FUNCTION_BLOCK FB_ProductionTank EXTENDS FB_SFC_Cycle IMPLEMENTS ITF_FB_SFC_Cycle
VAR_INPUT
	eElementID		: E_Element_List;
	
	stTankValves				:	st_TankValves		;
	stLineSourceValves			:	st_LineSourceValves	;
	stTriBlenderSourceValves	:	st_LineSourceValves	;
	stLineTargetValves			:	st_LineTargetValves	;
	stfbTriBlenderTargetValves	:	st_LineTargetValves	;

	
	
	//valOutlet		: E_Pis_Name;//Comment?
	//valLine			: E_Pis_Name;//Comment?
	//valTriBlender	: E_Pis_Name;//Comment?
	//valDrain		: E_Pis_Name;//Comment?
	//valCIP			: E_Pis_Name;//Comment?
	
	valFilling				: E_Pis_Name;
	valFillWater			: E_Pis_Name;
	valFillWaterDrain		: E_Pis_Name;
	valDrainTapWater		: E_Pis_Name;
	
	eTank_Name				: E_Tank_Name;

	
	sens_TankTemp			: E_ASense_Name	;//Tenk temperature sensor ID
	
	valCW_In				:	E_Pis_Name	;//Valve to control tank temperature In
	valCW_Out				:	E_Pis_Name	;//Valve to control tank temperature Out (always at 100 open)
	
	//pumpEnum			:	E_Pump_List	;
	
END_VAR
VAR_OUTPUT
END_VAR
VAR
	sTank_Name			: STRING;
	refElement			: REFERENCE TO FB_Element;
	refState_Long		: REFERENCE TO E_Element_State_Long;
	eReq				: E_Request_List;		
	eProcess			: E_Element_Process;
	eStatus				: E_Element_State_Long; // for HMI only as status
	
	fbPis				: FB_Piston;	
	
	//stPis_FillWater			: REFERENCE TO ST_Piston;
	//stPis_FillWaterDrain		: REFERENCE TO ST_Piston;
	//stPis_DrainTapWater		: REFERENCE TO ST_Piston;
	
	stPis_CWIn				: REFERENCE TO ST_Piston;
	stPis_CWOut				: REFERENCE TO ST_Piston;
	
	bTestingMode	:	BOOL	;//For testing purposes, to be deleted 
	bMoveStep		:	BOOL	;//For testing purposes, to be deleted 
	
	Call_TON	:	TON	;//Call ton for double request same object
	bTON_Active	:	BOOL	;
	
	// Temperature process control
	pc_TempCntrl	: REFERENCE TO FB_ProcessControl	;
	st_TempCntrl	: REFERENCE TO ST_ProcessControl	;
	bCntrlTemp		: BOOL	;
	bRunCIP			: BOOL	;
	
	ref_fbTankSensors			: REFERENCE TO FB_TankSensors;
	stTank_Level				: ST_Tank_Level;

	//888888888888888888888888888888888888888888
	stProdParam		: ST_Production_Parameter;
	//888888888888888888888888888888888888888888
	tonStirrer_time: TON;
	rTest: REAL := 16;
	bStirrerDirectionPositive: BOOL;
	
	delta_Tank_Volume		: REAL;
	memo_Tank_Level_start	: REAL;
	bRunOffline: BOOL;
	
	event_state_Update: INT;
	event_state_Update_sum: INT;
	event_state_Update_sum_last: INT;
	fbEvent_echo: FB_Event_echo;
	memo_Production_Storage_Mode: BOOL;
	memo_CIP_Pump_linked: BOOL;
	
	bStateUpdate_Available_HMI	: BOOL;

	
	
	fbFilling				: FB_Filling;		
	eFilling_State			: E_Filling_State;

END_VAR
VAR_IN_OUT

	fbTarget				: FB_Tank_Target;
	fbLineSource			: FB_Line_Source;
	fbLineTarget			: FB_Line_Target;
	fbTriBlenderSource		: FB_Line_Source;
	fbTriBlenderTarget		: FB_Line_Target;
	
	fbInterConnection_TriB	: FB_InterConnection;
	fbInterConnection_ProL	: FB_InterConnection;
	

	fb_PumpLine				: FB_Pump;
	fb_PumpTriBlender		: FB_Pump;
	fb_Stirrer				: FB_Pump;
END_VAR

act_GetReference();
act_Oper();
act_Call_Interface(); //There is no need to Call block if it comes from the outside
act_TempCntrl();
act_ExpirationTime();
act_Filling();

CASE eTank_Name OF
	E_Tank_Name.T1: sTank_Name:='Production Tank-T1';
	E_Tank_Name.T2: sTank_Name:='Production Tank-T2';
	E_Tank_Name.T3: sTank_Name:='Production Tank-T3';
	E_Tank_Name.T4: sTank_Name:='Production Tank-T4';
END_CASE

IF bTestingMode THEN;
	IF bMoveStep THEN;
		bMoveStep:=FALSE; 
	END_IF	
ELSE;
	bMoveStep:=TRUE; 
END_IF


IF stProdParam.bGetRecipe THEN;
	stProdParam.bGetRecipe:=FALSE;
	mGet_Recipe(indexRecipe:=stProdParam.hmiRecipeIndex+1);
END_IF
CASE eElementID	OF 
	E_Element_List.eTank_1,E_Element_List.eTank_2:;
		stProdParam.listRecipe:=g_Prod.listRecipe_Marinade;
	E_Element_List.eTank_3,E_Element_List.eTank_4:;
  		stProdParam.listRecipe:=g_Prod.listRecipe_Color;
END_CASE

stProdParam.timeRemainToStart:=mTimeRemainToStart();
stProdParam.timeProductionDuration:=mTimeProductionDuration();
refElement.ProdStatus:=stProdParam.eStatus;


IF refElement.m_Get_InterConnection()=E_InterConnection.NotConnected 
AND bReady
THEN;
	IF NOT bStateUpdate_Available_HMI THEN;
		refElement.fbEvent_echo.event();
		bStateUpdate_Available_HMI:=TRUE;
	END_IF	
ELSE; 
	IF bStateUpdate_Available_HMI THEN;
		refElement.fbEvent_echo.event();
		bStateUpdate_Available_HMI:=FALSE;
	END_IF
END_IF

m_Stirrer();
m_HMI();

ACTION _aCheck_Condition_Prod_End_active:
bStepDone:=FALSE;
IF fbInterConnection_ProL.bAvalableToDisconnect 
AND stProdParam.eStatus=E_Prod_Status.Active
THEN;
	bStepDone:=TRUE;
END_IF
END_ACTION

ACTION _aCheck_Condition_Product_active:
bStepDone:=FALSE;
IF fbInterConnection_ProL.bAvalableToConnect 
AND stProdParam.eStatus=E_Prod_Status.Active
THEN;
	bStepDone:=TRUE;
END_IF
END_ACTION

ACTION _aCheck_Condition_TriB_1_active_1:
bStepDone:=FALSE;
IF fbInterConnection_TriB.bAvalableToConnect
AND stProdParam.eStatus=E_Prod_Status.Active
AND m_Get_TriBlender_Clean()
THEN;
	bStepDone:=TRUE;
END_IF
END_ACTION

ACTION _aCheck_Condition_TriB_2_active:
bStepDone:=FALSE;
IF fbInterConnection_TriB.bAvalableToConnect 
AND stProdParam.eStatus=E_Prod_Status.Active
AND m_Get_TriBlender_Clean()
THEN;
	bStepDone:=TRUE;
END_IF
END_ACTION

ACTION _aClose_01_active:
bStepDone:=FALSE;
IF fbTarget.m_CheckStatus(eReqStatus:=E_Tank_Target.eClose) THEN;
	bStepDone:=TRUE;
END_IF
END_ACTION

ACTION _aClose_01_entry:
fbTarget.m_Run(eReqProc:=E_Tank_Target.eClose);
END_ACTION

ACTION _aClose_2_active:
bStepDone:=FALSE;
IF fbTarget.m_CheckStatus(eReqStatus:=E_Tank_Target.eClose) THEN;
	bStepDone:=TRUE;
END_IF
END_ACTION

ACTION _aClose_2_entry:
fbTarget.m_Run(eReqProc:=E_Tank_Target.eClose);
END_ACTION

ACTION _aClose_4_active:
bStepDone:=FALSE;
IF fbTarget.m_CheckStatus(eReqStatus:=E_Tank_Target.eClose) THEN;
	bStepDone:=TRUE;
END_IF
END_ACTION

ACTION _aClose_4_entry:
fbTarget.m_Run(eReqProc:=E_Tank_Target.eClose);
END_ACTION

ACTION _aClose_Drain_val_active:
//bStepDone:=FALSE;
IF fbTarget.m_CheckStatus(eReqStatus:=E_Tank_Target.eOpen) THEN;
(*ELSE
	fbTarget.m_Run(eReqProc:=E_Tank_Target.eOpen);*)
	bTON_Active:=TRUE;
END_IF
IF Call_TON.Q THEN
	bStepDone:=TRUE;
END_IF
END_ACTION

ACTION _aClose_Drain_val_entry:
bStepDone:=FALSE;
fbTarget.m_Run(eReqProc:=E_Tank_Target.eOpen);
bTON_Active:=FALSE;
END_ACTION

ACTION _aClose_Tank_active:
bStepDone:=FALSE;
IF fbTarget.m_CheckStatus(eReqStatus:=E_Tank_Target.eClose_DrainPipe) THEN;
	bStepDone:=TRUE;
END_IF
END_ACTION

ACTION _aClose_Tank_entry:
fbTarget.m_Run(eReqProc:=E_Tank_Target.eClose_DrainPipe);
END_ACTION

ACTION _aCollect_From_Prod_Line_active:
bStepDone:=FALSE;
delta_Tank_Volume:=ref_fbTankSensors.act_Volume-memo_Tank_Level_start;
IF FALSE 
OR delta_Tank_Volume>=stProdParam.stRecipe.Weight_to_Collect
OR Collect_From_Prod_Line.t>=T#40S
THEN;
	bStepDone:=TRUE;
END_IF
END_ACTION

ACTION _aCollect_From_TriB_Line_active:
bStepDone:=FALSE;
delta_Tank_Volume:=ref_fbTankSensors.act_Volume-memo_Tank_Level_start;
IF FALSE 
OR delta_Tank_Volume>=stProdParam.stRecipe.Weight_to_Collect
OR Collect_From_TriB_Line.t>=T#40S
THEN;
	bStepDone:=TRUE;
END_IF
END_ACTION

ACTION _aConn_Line_Source_TankA_active:
bStepDone:=FALSE;
IF fbLineSource.m_CheckStatus(eReqStatus:=E_Line_Source.eTank_A) THEN;
	bStepDone:=TRUE;
END_IF
END_ACTION

ACTION _aConn_Line_Source_TankA_entry:
fbLineSource.m_Run(eReqProc:=E_Line_Source.eTank_A);
END_ACTION

ACTION _aConn_Line_Source_TankB_active:
bStepDone:=FALSE;
IF fbLineSource.m_CheckStatus(eReqStatus:=E_Line_Source.eTank_B) THEN;
	bStepDone:=TRUE;
END_IF
END_ACTION

ACTION _aConn_Line_Source_TankB_entry:
fbLineSource.m_Run(eReqProc:=E_Line_Source.eTank_B);
END_ACTION

ACTION _aConn_Line_Target_TankA_active:
bStepDone:=FALSE;
IF fbLineTarget.m_CheckStatus(eReqStatus:=E_Line_Target.eTank_A) THEN;
	bTON_Active:=TRUE;
END_IF
IF Call_TON.Q THEN
	bStepDone:=TRUE;
END_IF
END_ACTION

ACTION _aConn_Line_Target_TankA_entry:
fbLineTarget.m_Run(eReqProc:=E_Line_Target.eTank_A);
bTON_Active:=FALSE;
END_ACTION

ACTION _aConn_Line_Target_TankB_active:
bStepDone:=FALSE;
IF fbLineTarget.m_CheckStatus(eReqStatus:=E_Line_Target.eTank_B) THEN;
	bTON_Active:=TRUE;
END_IF
IF Call_TON.Q THEN
	bStepDone:=TRUE;
END_IF
END_ACTION

ACTION _aConn_Line_Target_TankB_entry:
fbLineTarget.m_Run(eReqProc:=E_Line_Target.eTank_B);
bTON_Active:=FALSE;
END_ACTION

ACTION _aConn_Tank_active:
bStepDone:=FALSE;
IF fbTriBlenderSource.m_CheckStatus(eReqStatus:=E_Line_Source.eFillWater) 
//AND fbPis.m_CheckByRecipe(stPis:=stPis_FillWaterDrain, req:=E_Piston_Recipe_State.Release) 
THEN;
	bStepDone:=TRUE;
END_IF
END_ACTION

ACTION _aConn_Tank_entry:
fbTriBlenderSource.m_Run(eReqProc:=E_Line_Source.eFillWater);
//fbPis.m_SetByRecipe(stPis:=stPis_FillWaterDrain, req:=E_Piston_Recipe_State.Release);
END_ACTION

ACTION _aConn_Tri_Drain_active:
bStepDone:=FALSE;
IF fbTriBlenderTarget.m_CheckStatus(eReqStatus:=E_Line_Target.eDrain) THEN;
	bStepDone:=TRUE;
END_IF
END_ACTION

ACTION _aConn_Tri_Drain_entry:
fbTriBlenderTarget.m_Run(eReqProc:=E_Line_Target.eDrain);
END_ACTION

ACTION _aConn_Tri_TankA_2_active:
bStepDone:=FALSE;
IF fbTriBlenderSource.m_CheckStatus(eReqStatus:=E_Line_Source.eTank_A) THEN;
	bStepDone:=TRUE;
END_IF
END_ACTION

ACTION _aConn_Tri_TankA_2_entry:
fbTriBlenderSource.m_Run(eReqProc:=E_Line_Source.eTank_A);
END_ACTION

ACTION _aConn_Tri_TankB_2_active:
bStepDone:=FALSE;
IF fbTriBlenderSource.m_CheckStatus(eReqStatus:=E_Line_Source.eTank_B) THEN;
	bStepDone:=TRUE;
END_IF
END_ACTION

ACTION _aConn_Tri_TankB_2_entry:
fbTriBlenderSource.m_Run(eReqProc:=E_Line_Source.eTank_B);
END_ACTION

ACTION _aConn_Tri_TapWater_active:
bStepDone:=FALSE;
IF fbTriBlenderSource.m_CheckStatus(eReqStatus:=E_Line_Source.eTapWater) 
//AND fbPis.m_CheckByRecipe(stPis:=stPis_DrainTapWater, req:=E_Piston_Recipe_State.Release) 
THEN;
	bTON_Active:=TRUE;
END_IF
IF Call_TON.Q THEN
	bStepDone:=TRUE;
END_IF
END_ACTION

ACTION _aConn_Tri_TapWater_entry:
fbTriBlenderSource.m_Run(eReqProc:=E_Line_Source.eTapWater);
//fbPis.m_SetByRecipe(stPis:=stPis_DrainTapWater, req:=E_Piston_Recipe_State.Release);
bTON_Active:=FALSE;
END_ACTION

ACTION _aConn_Tri_ToTankA_1_active:
bStepDone:=FALSE;
IF fbTriBlenderTarget.m_CheckStatus(eReqStatus:=E_Line_Target.eTank_A) THEN;
	bStepDone:=TRUE;
END_IF
END_ACTION

ACTION _aConn_Tri_ToTankA_1_entry:
fbTriBlenderTarget.m_Run(eReqProc:=E_Line_Target.eTank_A);
END_ACTION

ACTION _aConn_Tri_ToTankA_2_active:
bStepDone:=FALSE;
IF fbTriBlenderTarget.m_CheckStatus(eReqStatus:=E_Line_Target.eTank_A) THEN;
	bStepDone:=TRUE;
END_IF
END_ACTION

ACTION _aConn_Tri_ToTankA_2_entry:
fbTriBlenderTarget.m_Run(eReqProc:=E_Line_Target.eTank_A);
END_ACTION

ACTION _aConn_Tri_ToTankB_1_active:
bStepDone:=FALSE;
IF fbTriBlenderTarget.m_CheckStatus(eReqStatus:=E_Line_Target.eTank_B) THEN;
	bStepDone:=TRUE;
END_IF
END_ACTION

ACTION _aConn_Tri_ToTankB_1_entry:
fbTriBlenderTarget.m_Run(eReqProc:=E_Line_Target.eTank_B);
END_ACTION

ACTION _aConn_Tri_ToTankB_2_active:
bStepDone:=FALSE;
IF fbTriBlenderTarget.m_CheckStatus(eReqStatus:=E_Line_Target.eTank_B) THEN;
	bStepDone:=TRUE;
END_IF
END_ACTION

ACTION _aConn_Tri_ToTankB_2_entry:
fbTriBlenderTarget.m_Run(eReqProc:=E_Line_Target.eTank_B);
END_ACTION

ACTION _aConn_TriB_Color_active_1:
bStepDone:=FALSE;
IF fbTriBlender_Select.m_CheckStatus(eReqStatus:=E_TriBlenderSelect.eColor) THEN;
	bStepDone:=TRUE;
END_IF
END_ACTION

ACTION _aConn_TriB_Color_entry_1:
fbTriBlender_Select.m_Set_Request(eSetReg:=E_TriBlenderSelect.eColor);
END_ACTION

ACTION _aConn_TriB_Marinade_active_1:
bStepDone:=FALSE;
IF fbTriBlender_Select.m_CheckStatus(eReqStatus:=E_TriBlenderSelect.eMarinade) THEN;
	bStepDone:=TRUE;
END_IF
END_ACTION

ACTION _aConn_TriB_Marinade_entry_1:
fbTriBlender_Select.m_Set_Request(eSetReg:=E_TriBlenderSelect.eMarinade);
END_ACTION

ACTION _aDis_Conn_Tank_active:
bStepDone:=FALSE;
IF fbTriBlenderSource.m_CheckStatus(eReqStatus:=E_Line_Source.eClose) 
AND fbTriBlenderTarget.m_CheckStatus(eReqStatus:=E_Line_Target.eDrain) 
THEN;
	bStepDone:=TRUE;
END_IF
END_ACTION

ACTION _aDis_Conn_Tank_entry:
fbTriBlenderSource.m_Run(eReqProc:=E_Line_Source.eClose);
fbTriBlenderTarget.m_Run(eReqProc:=E_Line_Target.eDrain);
END_ACTION

ACTION _aDisconn_Tri_Tank_active:
bStepDone:=FALSE;
IF fbTriBlenderSource.m_CheckStatus(eReqStatus:=E_Line_Source.eClose) THEN;
	bTON_Active:=TRUE;
END_IF
IF Call_TON.Q THEN
	bStepDone:=TRUE;
END_IF
END_ACTION

ACTION _aDisconn_Tri_Tank_entry:
fbTriBlenderSource.m_Run(eReqProc:=E_Line_Source.eClose);
bTON_Active:=FALSE;
END_ACTION

ACTION _aDisconnect_TapWater_02_active:
bStepDone:=FALSE;
IF fbTriBlenderSource.m_CheckStatus(eReqStatus:=E_Line_Source.eDrain) THEN;
	bStepDone:=TRUE;
END_IF
END_ACTION

ACTION _aDisconnect_TapWater_02_entry:
fbTriBlenderSource.m_Run(eReqProc:=E_Line_Source.eDrain);
END_ACTION

ACTION _aDissolving_entry:
bDisolvingProcess_Done:=FALSE;
bDisolvingProcess_Active:=FALSE;
END_ACTION

ACTION _aDissolving_Proc_active:
bStepDone:=FALSE;

IF bDisolvingProcess_Done 
//AND fbDissolving.bD
THEN;
	
END_IF
END_ACTION

ACTION _aDissolving_Proc_entry:

bDisolvingProcess_Active:=TRUE;
fbDissolving.mRun();
END_ACTION

ACTION _aDissolving_Proc_exit:
bDisolvingProcess_Done:=FALSE;
bDisolvingProcess_Active:=FALSE;
END_ACTION

ACTION _aDone_entry:
eProcess:=E_Element_Process.eNone;
eReq:=E_Request_List.eNone;
bRun:=FALSE;
bDone:=TRUE;
END_ACTION

ACTION _aDrain_All_Marinade_Lines_active:
bStepDone:=FALSE;
IF TRUE
//AND fbTarget.m_CheckStatus(eReqStatus:=E_Tank_Target.eClose_DrainPipe) 
AND fbTriBlenderSource.m_CheckStatus(eReqStatus:=E_Line_Source.eDrain)
AND fbTriBlenderTarget.m_CheckStatus(eReqStatus:=E_Line_Target.eDrain)
AND fbTriBlender_Select.m_CheckStatus(eReqStatus:=E_TriBlenderSelect.eDrain)
AND TRUE
AND TRUE
THEN;
	bStepDone:=TRUE;
END_IF
END_ACTION

ACTION _aDrain_All_Marinade_Lines_entry:
//fbTarget.m_Run(eReqProc:=E_Tank_Target.eClose_DrainPipe);
fbTriBlenderSource.m_Run(eReqProc:=E_Line_Source.eDrain);
fbTriBlenderTarget.m_Run(eReqProc:=E_Line_Target.eDrain);
fbTriBlender_Select.m_Set_Request(eSetReg:=E_TriBlenderSelect.eDrain);
END_ACTION

ACTION _aDrain_Pipe_active:
bStepDone:=FALSE;
IF fbTarget.m_CheckStatus(eReqStatus:=E_Tank_Target.eClose_DrainPipe) THEN;
	bTON_Active:=TRUE;
END_IF
IF Call_TON.Q THEN
	bStepDone:=TRUE;
END_IF
END_ACTION

ACTION _aDrain_Pipe_Close_active:
bStepDone:=FALSE;
IF fbTarget.m_CheckStatus(eReqStatus:=E_Tank_Target.eClose) THEN;
	bStepDone:=TRUE;
END_IF
END_ACTION

ACTION _aDrain_Pipe_Close_entry:
fbTarget.m_Run(eReqProc:=E_Tank_Target.eClose);
END_ACTION

ACTION _aDrain_Pipe_entry:
fbTarget.m_Run(eReqProc:=E_Tank_Target.eClose_DrainPipe);
bTON_Active:=FALSE;
END_ACTION

ACTION _aDrain_Production_Line_active:
bStepDone:=FALSE;
IF TRUE
AND fbTarget.m_CheckStatus(eReqStatus:=E_Tank_Target.eClose_DrainPipe) 
AND fbLineSource.m_CheckStatus(eReqStatus:=E_Line_Source.eDrain)
AND fbLineTarget.m_CheckStatus(eReqStatus:=E_Line_Target.eDrain)
AND TRUE
THEN;
	bStepDone:=TRUE;
END_IF
END_ACTION

ACTION _aDrain_Production_Line_entry:
fbTarget.m_Run(eReqProc:=E_Tank_Target.eClose_DrainPipe);
fbLineSource.m_Run(eReqProc:=E_Line_Source.eDrain);
fbLineTarget.m_Run(eReqProc:=E_Line_Target.eDrain);
END_ACTION

ACTION _aDrain_Tri_Line_active:
bStepDone:=FALSE;
IF fbTriBlenderTarget.m_CheckStatus(eReqStatus:=E_Line_Target.eDrain) THEN;
	bStepDone:=TRUE;
END_IF
END_ACTION

ACTION _aDrain_Tri_Line_entry:
fbTriBlenderTarget.m_Run(eReqProc:=E_Line_Target.eDrain);
END_ACTION

ACTION _aDrain_Tri_ToDrain_active:
bStepDone:=FALSE;
IF fbTriBlenderTarget.m_CheckStatus(eReqStatus:=E_Line_Target.eDrain) THEN;
	bTON_Active:=TRUE;
END_IF
IF Call_TON.Q THEN
	bStepDone:=TRUE;
END_IF

(*
delta_Tank_Volume:=ref_fbTankSensors.act_Volume-memo_Tank_Level_start;
IF bStepDone
AND  
AND (delta_Tank_Volume>=stProdParam.stRecipe.Weight_to_Drain
	OR Drain_Tri_ToDrain.t>=T#30S)
THEN;
	//bStepDone:=TRUE;
ELSE;
	bStepDone:=FALSE;
END_IF
*)
END_ACTION

ACTION _aDrain_Tri_ToDrain_entry:
fbTriBlenderTarget.m_Run(eReqProc:=E_Line_Target.eDrain);
bTON_Active:=FALSE;
END_ACTION

ACTION _aDrain_Tri_ToTankA_active:
bStepDone:=FALSE;
IF fbTriBlenderTarget.m_CheckStatus(eReqStatus:=E_Line_Target.eTank_A) THEN;
	bTON_Active:=TRUE;
END_IF
IF Call_TON.Q THEN
	bStepDone:=TRUE;
END_IF
END_ACTION

ACTION _aDrain_Tri_ToTankA_entry:
fbTriBlenderTarget.m_Run(eReqProc:=E_Line_Target.eTank_A);
bTON_Active:=FALSE;
END_ACTION

ACTION _aDrain_Tri_ToTankB_active:
bStepDone:=FALSE;
IF fbTriBlenderTarget.m_CheckStatus(eReqStatus:=E_Line_Target.eTank_B) THEN;
	bTON_Active:=TRUE;
END_IF
IF Call_TON.Q THEN
	bStepDone:=TRUE;
END_IF
END_ACTION

ACTION _aDrain_Tri_ToTankB_entry:
fbTriBlenderTarget.m_Run(eReqProc:=E_Line_Target.eTank_B);
bTON_Active:=FALSE;
END_ACTION

ACTION _aDrain_Trib_Line_01_active:
bStepDone:=FALSE;
IF fbTriBlender_Select.m_CheckStatus(eReqStatus:=E_TriBlenderSelect.eDrain) THEN;
	bStepDone:=TRUE;
END_IF
END_ACTION

ACTION _aDrain_Trib_Line_01_entry:
fbTriBlender_Select.m_Set_Request(eSetReg:=E_TriBlenderSelect.eDrain);
END_ACTION

ACTION _aDrain_Trib_Line_02_active:
bStepDone:=FALSE;
IF fbTriBlender_Select.m_CheckStatus(eReqStatus:=E_TriBlenderSelect.eDrain)
OR fbTriBlender_Select.m_CheckStatus(eReqStatus:=E_TriBlenderSelect.eMarinade) THEN;//marinade =>> drain time finish
	bStepDone:=TRUE;
END_IF
END_ACTION

ACTION _aDrain_Trib_Line_02_entry:
fbTriBlender_Select.m_Set_Request(eSetReg:=E_TriBlenderSelect.eDrain);
END_ACTION

ACTION _aDraining_Time_active:
bStepDone:=FALSE;
IF stTank_Level.e_state=E_Tank_Level.eEmpty THEN;
	bStepDone:=TRUE;
END_IF
END_ACTION

ACTION _aDrainOpen_01_active:
bStepDone:=FALSE;
IF fbTarget.m_CheckStatus(eReqStatus:=E_Tank_Target.eDrain) THEN;
	bStepDone:=TRUE;
END_IF
END_ACTION

ACTION _aDrainOpen_01_entry:
fbTarget.m_Run(eReqProc:=E_Tank_Target.eDrain);
END_ACTION

ACTION _aDriin_Tank_active:
bStepDone:=FALSE;
IF stTank_Level.e_state=E_Tank_Level.eEmpty THEN;
	bStepDone:=TRUE;
END_IF
END_ACTION

ACTION _aDriin_Tank_entry:
fbTarget.m_Run(eReqProc:=E_Tank_Target.eDrain);
END_ACTION

ACTION _aInit_Base_active:
bStepDone:=FALSE;
IF TRUE
AND refState_Long<>E_Element_State_Long.eProduction
AND fbTarget.m_CheckStatus(eReqStatus:=E_Tank_Target.eClose_DrainPipe) 
AND TRUE
THEN;
	bStepDone:=TRUE;
ELSIF refState_Long=E_Element_State_Long.eProduction THEN;
	bStepDone:=TRUE;
END_IF
END_ACTION

ACTION _aInit_Base_entry:
IF refState_Long<>E_Element_State_Long.eProduction THEN;	
	fb_PumpLine.m_Stop();
	fbTarget.m_Run(eReqProc:=E_Tank_Target.eClose_DrainPipe);
END_IF
END_ACTION

ACTION _aInit_Production_Line_active:
bStepDone:=FALSE;
IF TRUE
AND refState_Long<>E_Element_State_Long.eProduction
AND fbTarget.m_CheckStatus(eReqStatus:=E_Tank_Target.eClose_DrainPipe) 
AND fbLineSource.m_CheckStatus(eReqStatus:=E_Line_Source.eDrain)
AND fbLineTarget.m_CheckStatus(eReqStatus:=E_Line_Target.eDrain)
AND (NOT fbInterConnection_ProL.bActive)
AND TRUE
THEN;
	bStepDone:=TRUE;
ELSIF refState_Long=E_Element_State_Long.eProduction THEN;
	bStepDone:=TRUE;
END_IF
END_ACTION

ACTION _aInit_Production_Line_entry:
IF refState_Long<>E_Element_State_Long.eProduction THEN;	
	fb_PumpLine.m_Stop();
	fbTarget.m_Run(eReqProc:=E_Tank_Target.eClose_DrainPipe);
	fbLineSource.m_Run(eReqProc:=E_Line_Source.eDrain);
	fbLineTarget.m_Run(eReqProc:=E_Line_Target.eDrain);
	fbInterConnection_ProL.reqDisconnect:=TRUE;
END_IF
END_ACTION

ACTION _aInit_Tank_active:
SFCReset:=FALSE;
END_ACTION

ACTION _aInit_Tank_exit:
IF eProcess=E_Element_Process.eFill_Water THEN;
	mClearProduction(state:=E_Element_State_Long.eOff);
END_IF

eProcess:=E_Element_Process.eNone;
eReq:=E_Request_List.eNone;
memo_Production_Storage_Mode:=FALSE;
END_ACTION

ACTION _aInit_TriBlender_Line_active:
bStepDone:=FALSE;
IF TRUE
AND fbTarget.m_CheckStatus(eReqStatus:=E_Tank_Target.eClose_DrainPipe) 
AND fbTriBlenderSource.m_CheckStatus(eReqStatus:=E_Line_Source.eDrain)
AND fbTriBlenderTarget.m_CheckStatus(eReqStatus:=E_Line_Target.eDrain)
AND fbTriBlender_Select.m_CheckStatus(eReqStatus:=E_TriBlenderSelect.eDrain)
AND (NOT fbInterConnection_TriB.bActive)
AND TRUE
THEN;
	bStepDone:=TRUE;
END_IF
END_ACTION

ACTION _aInit_TriBlender_Line_entry:
fb_PumpTriBlender.m_Stop();
fbTarget.m_Run(eReqProc:=E_Tank_Target.eClose_DrainPipe);
fbTriBlenderSource.m_Run(eReqProc:=E_Line_Source.eDrain);
fbTriBlenderTarget.m_Run(eReqProc:=E_Line_Target.eDrain);
fbTriBlender_Select.m_Set_Request(eSetReg:=E_TriBlenderSelect.eDrain);
fbInterConnection_TriB.reqDisconnect:=TRUE;
fbDissolving.mResetCycle();
END_ACTION

ACTION _aInterConnect_Prod_active:
bStepDone:=FALSE;
IF fbInterConnection_ProL.bActive THEN;
	bStepDone:=TRUE;
END_IF
END_ACTION

ACTION _aInterConnect_Prod_Dis_active:
bStepDone:=FALSE;
IF NOT fbInterConnection_ProL.bActive THEN;
	bStepDone:=TRUE;
END_IF
END_ACTION

ACTION _aInterConnect_Prod_Dis_entry:
fbInterConnection_ProL.reqDisconnect:=TRUE;
END_ACTION

ACTION _aInterConnect_Prod_entry:
fbInterConnection_ProL.reqConnect:=TRUE;

IF trn_Tank_Marinade THEN;
	//fbElement[E_Element_List.eTriBlender_Marinada].m_Set_Dissolveng_active_memo();
ELSIF trn_Tank_Color THEN;
	//fbElement[E_Element_List.eTriBlender_Color].m_Set_Dissolveng_active_memo();
END_IF
END_ACTION

ACTION _aInterConnect_TriB_1_active:
bStepDone:=FALSE;
IF fbInterConnection_TriB.bActive THEN;
	bStepDone:=TRUE;
END_IF
END_ACTION

ACTION _aInterConnect_TriB_1_entry:
fbInterConnection_TriB.reqConnect:=TRUE;
END_ACTION

ACTION _aInterConnect_TriB_2_active:
bStepDone:=FALSE;
IF fbInterConnection_TriB.bActive THEN;
	bStepDone:=TRUE;
	
	refElement.m_Set_Dissolveng_active_memo();
	IF trn_Tank_Marinade THEN;
		fbElement[E_Element_List.eTriBlender_Marinada].m_Set_Dissolveng_active_memo();
	ELSIF trn_Tank_Color THEN;
		fbElement[E_Element_List.eTriBlender_Color].m_Set_Dissolveng_active_memo();
	ELSE;
		bStepDone:=FALSE;
	END_IF	
	
END_IF
END_ACTION

ACTION _aInterConnect_TriB_2_entry:
fbInterConnection_TriB.reqConnect:=TRUE;
END_ACTION

ACTION _aInterConnect_TriB_Dis_1_active:
bStepDone:=FALSE;
IF NOT fbInterConnection_TriB.bActive THEN;
	bStepDone:=TRUE;
END_IF
END_ACTION

ACTION _aInterConnect_TriB_Dis_1_entry:
fbInterConnection_TriB.reqDisconnect:=TRUE;
END_ACTION

ACTION _aInterConnect_TriB_Dis_2_active:
bStepDone:=FALSE;
IF NOT fbInterConnection_TriB.bActive THEN;
	bStepDone:=TRUE;
END_IF
END_ACTION

ACTION _aInterConnect_TriB_Dis_2_entry:
fbInterConnection_TriB.reqDisconnect:=TRUE;
END_ACTION

ACTION _aLineSource_Close_active:
bStepDone:=FALSE;
IF fbLineSource.m_CheckStatus(eReqStatus:=E_Line_Source.eClose) 
THEN;
	bStepDone:=TRUE;
END_IF
END_ACTION

ACTION _aLineSource_Close_entry:
fbLineSource.m_Run(eReqProc:=E_Line_Source.eClose);
END_ACTION

ACTION _aLineSource_TapWater_active:
bStepDone:=FALSE;
IF fbLineSource.m_CheckStatus(eReqStatus:=E_Line_Source.eTapWater) 
THEN;
	bStepDone:=TRUE;
END_IF
END_ACTION

ACTION _aLineSource_TapWater_entry:
fbLineSource.m_Run(eReqProc:=E_Line_Source.eTapWater);
bTON_Active:=FALSE;
END_ACTION

ACTION _aLineTarget_Drain_1_active:
bStepDone:=FALSE;
IF fbLineTarget.m_CheckStatus(eReqStatus:=E_Line_Target.eDrain) THEN;
	bStepDone:=TRUE;
END_IF
END_ACTION

ACTION _aLineTarget_Drain_1_entry:
fbLineTarget.m_Run(eReqProc:=E_Line_Target.eDrain);
END_ACTION

ACTION _aLineTarget_Drain_2_active:
bStepDone:=FALSE;
IF fbLineTarget.m_CheckStatus(eReqStatus:=E_Line_Target.eDrain) THEN;
	bTON_Active:=TRUE;
END_IF
IF Call_TON.Q THEN
	bStepDone:=TRUE;
END_IF
END_ACTION

ACTION _aLineTarget_Drain_2_entry:
fbLineTarget.m_Run(eReqProc:=E_Line_Target.eDrain);
bTON_Active:=FALSE;
END_ACTION

ACTION _aLineTarget_TankA_active:
bStepDone:=FALSE;
IF fbLineTarget.m_CheckStatus(eReqStatus:=E_Line_Target.eTank_A) THEN;
	bTON_Active:=TRUE;
END_IF
IF Call_TON.Q THEN
	bStepDone:=TRUE;
END_IF
END_ACTION

ACTION _aLineTarget_TankA_entry:
fbLineTarget.m_Run(eReqProc:=E_Line_Target.eTank_A);
bTON_Active:=FALSE;
END_ACTION

ACTION _aLineTarget_TankB_active:
bStepDone:=FALSE;
IF fbLineTarget.m_CheckStatus(eReqStatus:=E_Line_Target.eTank_B) THEN;
	bTON_Active:=TRUE;
END_IF
IF Call_TON.Q THEN
	bStepDone:=TRUE;
END_IF
END_ACTION

ACTION _aLineTarget_TankB_entry:
fbLineTarget.m_Run(eReqProc:=E_Line_Target.eTank_B);
bTON_Active:=FALSE;
END_ACTION

ACTION _aOpen_Drain_Pipe_active:
bStepDone:=FALSE;
IF fbTarget.m_CheckStatus(eReqStatus:=E_Tank_Target.eClose_DrainPipe) THEN;
	bStepDone:=TRUE;
END_IF
END_ACTION

ACTION _aOpen_Drain_Pipe_entry:
fbTarget.m_Run(eReqProc:=E_Tank_Target.eClose_DrainPipe);
END_ACTION

ACTION _aPumpLine_Auto_1_entry:
//fb_PumpLine.m_Auto();
END_ACTION

ACTION _aPumpLine_Start_1_active:

END_ACTION

ACTION _aPumpLine_Start_1_entry:
fb_PumpLine.m_Run(RPM:=stProdParam.stRecipe.FlowRate_Production);
END_ACTION

ACTION _aPumpLine_Start_2_entry:
fb_PumpLine.m_Run(RPM:=stProdParam.stRecipe.FlowRate_Production);
memo_Tank_Level_start:=ref_fbTankSensors.act_Volume;
END_ACTION

ACTION _aPumpLine_Stop_1_entry:
fb_PumpLine.m_Stop();
END_ACTION

ACTION _aPumpLine_Stop_2_entry:

IF trn_Tank_Marinade THEN;
	fb_PumpLine.m_Stop();
END_IF
END_ACTION

ACTION _aPumpLine_Stop_3_entry:
fb_PumpLine.m_Stop();
END_ACTION

ACTION _aPumpLine_Stop_4_entry:
fb_PumpLine.m_Stop();
END_ACTION

ACTION _aReady_active:


CASE refElement.eState_Long OF
	E_Element_State_Long.eOff,E_Element_State_Long.eStandby:;
			IF eReq=E_Request_List.eDrain THEN;
				eProcess:=E_Element_Process.eDrain;
			END_IF

	E_Element_State_Long.eCIP_5_Done:;
			IF eReq=E_Request_List.eWaterPrepare THEN;
				eProcess:=E_Element_Process.eFill_Water;
			END_IF	
			
	E_Element_State_Long.eWaterReady:;
			IF eReq=E_Request_List.eDissolve THEN;
				eProcess:=E_Element_Process.eDissolving;
			END_IF	
			IF eReq=E_Request_List.eFinish THEN;
				mClearProduction(state:=E_Element_State_Long.eStandby);
			END_IF
	E_Element_State_Long.eReady:;
			IF eReq=E_Request_List.eProduction THEN;
				eProcess:=E_Element_Process.eConnectionToLine;
			END_IF	
			IF eReq=E_Request_List.eFinish THEN;
				mClearProduction(state:=E_Element_State_Long.eStandby);
			END_IF			

	E_Element_State_Long.eProduction:;
			IF eReq=E_Request_List.eDisconnectTank THEN;
				eProcess:=E_Element_Process.eDisconnection;
			END_IF	
			
			IF fbInterConnection_ProL.bAvalableToDisconnect 
			AND m_Production_Run_Pump()
			THEN;
				IF memo_Production_Storage_Mode THEN;
					fb_PumpLine.m_Run(RPM:=stProdParam.stRecipe.FlowRate_Storage);
				ELSE;
					fb_PumpLine.m_Run(RPM:=stProdParam.stRecipe.FlowRate_Production);
				END_IF
				
			ELSE;
				fb_PumpLine.m_Stop();
			END_IF		

	E_Element_State_Long.eEmpty:;
			IF eReq=E_Request_List.eFinish THEN;
				mClearProduction(state:=E_Element_State_Long.eStandby);
			END_IF	

	E_Element_State_Long.eExpired:;
		CASE refElement.eState_Long_Expiered OF
			
			E_Element_State_Long.eProduction:;	
				IF eReq=E_Request_List.eDisconnectTank THEN;
					eProcess:=E_Element_Process.eDisconnection;
				END_IF
				
				IF fbInterConnection_ProL.bAvalableToDisconnect 
				AND m_Production_Run_Pump()
				THEN;
					IF memo_Production_Storage_Mode THEN;
						fb_PumpLine.m_Run(RPM:=stProdParam.stRecipe.FlowRate_Storage);
					ELSE;
						fb_PumpLine.m_Run(RPM:=stProdParam.stRecipe.FlowRate_Production);
					END_IF
					
				ELSE;
					fb_PumpLine.m_Stop();
				END_IF	
		ELSE
			IF eReq=E_Request_List.eFinish THEN;
				mClearProduction(state:=E_Element_State_Long.eStandby);
			END_IF			
		END_CASE
		
END_CASE
END_ACTION

ACTION _aReady_entry:

END_ACTION

ACTION _aReady_exit:
bRun:=TRUE;
bDone:=FALSE;
//bCntrlTemp:=TRUE;
END_ACTION

ACTION _aStart_TriPump_1_active:
bStepDone:=TRUE;
END_ACTION

ACTION _aStart_TriPump_1_entry:
fb_PumpTriBlender.m_Run(RPM:=stProdParam.stRecipe.FlowRate_WaterPushing);
END_ACTION

ACTION _aStart_TriPump_2_active:
bStepDone:=TRUE;
END_ACTION

ACTION _aStart_TriPump_2_entry:
fb_PumpTriBlender.m_Run(RPM:=stProdParam.stRecipe.FlowRate_WaterPushing);
END_ACTION

ACTION _aStart_TriPump_3_active:
bStepDone:=TRUE;
END_ACTION

ACTION _aStart_TriPump_3_entry:
fb_PumpTriBlender.m_Run(RPM:=stProdParam.stRecipe.FlowRate_WaterPushing);
memo_Tank_Level_start:=ref_fbTankSensors.act_Volume;
END_ACTION

ACTION _aState_Update_01_entry:
refState_Long:=E_Element_State_Long.eNotClean;
END_ACTION

ACTION _aState_Update_02_entry:
refState_Long:=E_Element_State_Long.eWaterReady;
END_ACTION

ACTION _aState_Update_03_entry:
refState_Long:=E_Element_State_Long.eReady;
END_ACTION

ACTION _aState_Update_04_entry:
refState_Long:=E_Element_State_Long.eProduction;
END_ACTION

ACTION _aState_Update_05_entry:
refState_Long:=E_Element_State_Long.eReady;
END_ACTION

ACTION _aStop_TriPump_1_active:
bStepDone:=TRUE;
END_ACTION

ACTION _aStop_TriPump_1_entry:
fb_PumpTriBlender.m_Stop();
END_ACTION

ACTION _aStop_TriPump_2_active:
bStepDone:=TRUE;
END_ACTION

ACTION _aStop_TriPump_2_entry:
fb_PumpTriBlender.m_Stop();
END_ACTION

ACTION _aStop_TriPump_3_active:
bStepDone:=TRUE;
END_ACTION

ACTION _aStop_TriPump_3_entry:
fb_PumpTriBlender.m_Stop();
END_ACTION

ACTION _aTank_Drain_active:
bStepDone:=FALSE;
IF fbTarget.m_CheckStatus(eReqStatus:=E_Tank_Target.eDrain) THEN;
	bTON_Active:=TRUE;
	
ELSIF Tank_Drain.t>=T#3S THEN; // max time to detect drain open
	bStepDone:=TRUE;
END_IF
IF Call_TON.Q THEN
	bStepDone:=TRUE;
END_IF
END_ACTION

ACTION _aTank_Drain_entry:
fbTarget.m_Run(eReqProc:=E_Tank_Target.eDrain);
bTON_Active:=FALSE;
END_ACTION

ACTION _aTank_Open_active:
bStepDone:=FALSE;
IF fbTarget.m_CheckStatus(eReqStatus:=E_Tank_Target.eOpen) THEN;
	bTON_Active:=TRUE;
END_IF
IF Call_TON.Q THEN
	bStepDone:=TRUE;
END_IF
END_ACTION

ACTION _aTank_Open_entry:
fbTarget.m_Run(eReqProc:=E_Tank_Target.eOpen);
bTON_Active:=FALSE;
END_ACTION

ACTION _aWater_Fill_active:
bStepDone:=FALSE;
IF TRUE 
AND TRUE//Reserved for tank level from recipe
//AND ref_fbTankSensors.get_stTankLevel().rTankLevel>=stProdParam.stRecipe.arr_Component[1].rWeight
AND fbTarget.stTankLevel.rTankLevel>=stProdParam.stRecipe.arr_Component[1].rWeight
THEN;
	bStepDone:=TRUE;
	
//temp overweight protection
ELSIF stT3_Sens.rTankLevel+stT4_Sens.rTankLevel>1000 THEN;
	bStepDone:=TRUE;
	
ELSIF bRunOffline 
AND Water_Fill.t>=T#10S
THEN
	bStepDone:=TRUE;
END_IF
END_ACTION

ACTION act_Call_Interface:
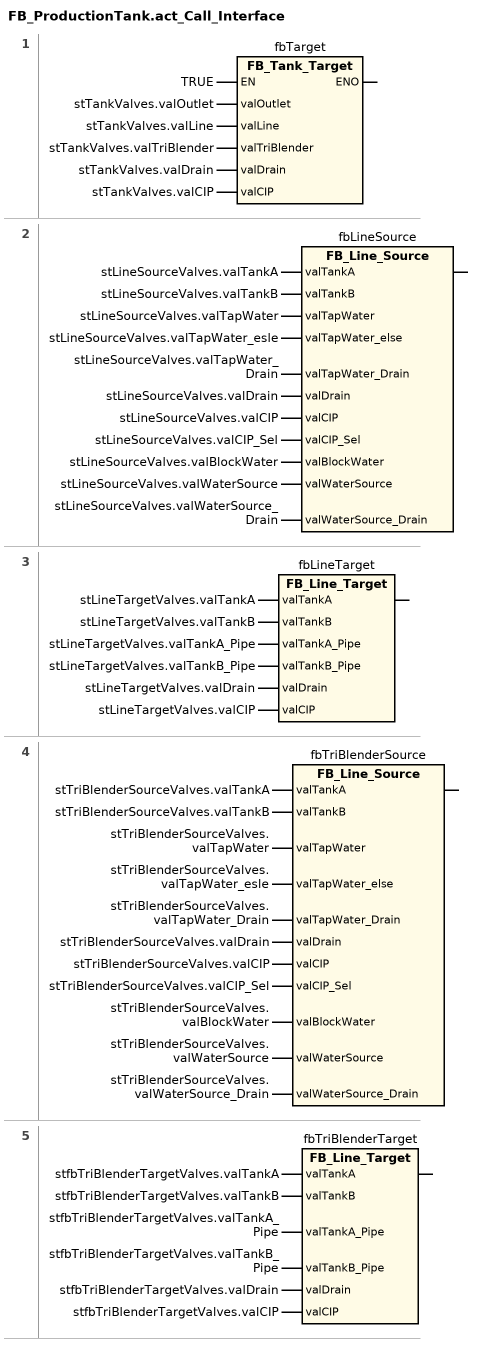
// NETWORK 1
fbTarget(
    valOutlet := stTankValves.valOutlet,
    valLine := stTankValves.valLine,
    valTriBlender := stTankValves.valTriBlender,
    valDrain := stTankValves.valDrain,
    valCIP := stTankValves.valCIP); // FB_Tank_Target

// NETWORK 2
fbLineSource(
    valTankA := stLineSourceValves.valTankA,
    valTankB := stLineSourceValves.valTankB,
    valTapWater := stLineSourceValves.valTapWater,
    valTapWater_else := stLineSourceValves.valTapWater_esle,
    valTapWater_Drain := stLineSourceValves.valTapWater_Drain,
    valDrain := stLineSourceValves.valDrain,
    valCIP := stLineSourceValves.valCIP,
    valCIP_Sel := stLineSourceValves.valCIP_Sel,
    valBlockWater := stLineSourceValves.valBlockWater,
    valWaterSource := stLineSourceValves.valWaterSource,
    valWaterSource_Drain := stLineSourceValves.valWaterSource_Drain); // FB_Line_Source

// NETWORK 3
fbLineTarget(
    valTankA := stLineTargetValves.valTankA,
    valTankB := stLineTargetValves.valTankB,
    valTankA_Pipe := stLineTargetValves.valTankA_Pipe,
    valTankB_Pipe := stLineTargetValves.valTankB_Pipe,
    valDrain := stLineTargetValves.valDrain,
    valCIP := stLineTargetValves.valCIP); // FB_Line_Target

// NETWORK 4
fbTriBlenderSource(
    valTankA := stTriBlenderSourceValves.valTankA,
    valTankB := stTriBlenderSourceValves.valTankB,
    valTapWater := stTriBlenderSourceValves.valTapWater,
    valTapWater_else := stTriBlenderSourceValves.valTapWater_esle,
    valTapWater_Drain := stTriBlenderSourceValves.valTapWater_Drain,
    valDrain := stTriBlenderSourceValves.valDrain,
    valCIP := stTriBlenderSourceValves.valCIP,
    valCIP_Sel := stTriBlenderSourceValves.valCIP_Sel,
    valBlockWater := stTriBlenderSourceValves.valBlockWater,
    valWaterSource := stTriBlenderSourceValves.valWaterSource,
    valWaterSource_Drain := stTriBlenderSourceValves.valWaterSource_Drain); // FB_Line_Source

// NETWORK 5
fbTriBlenderTarget(
    valTankA := stfbTriBlenderTargetValves.valTankA,
    valTankB := stfbTriBlenderTargetValves.valTankB,
    valTankA_Pipe := stfbTriBlenderTargetValves.valTankA_Pipe,
    valTankB_Pipe := stfbTriBlenderTargetValves.valTankB_Pipe,
    valDrain := stfbTriBlenderTargetValves.valDrain,
    valCIP := stfbTriBlenderTargetValves.valCIP); // FB_Line_Target

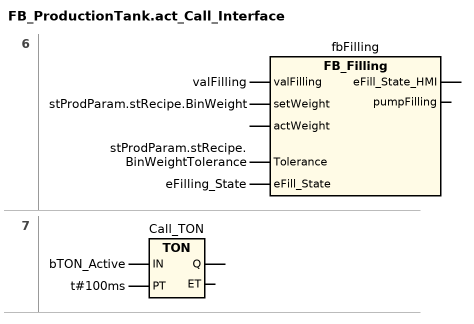
// NETWORK 6
fbFilling(
    valFilling := valFilling,
    setWeight := stProdParam.stRecipe.BinWeight,
    Tolerance := stProdParam.stRecipe.BinWeightTolerance,
    eFill_State := eFilling_State); // FB_Filling

// NETWORK 7
Call_TON(IN := bTON_Active, PT := t#100ms); // TON
END_ACTION

ACTION act_ExpirationTime:
IF stProdParam.eStatus=E_Prod_Status.Active 
THEN;
	refElement.m_Set_ExpirationDuration(eExTime_set:=E_ExTime.eProduct, setTime:=stProdParam.stRecipe.ExpirationTime);
	refElement.m_Set_ExpirationDuration(eExTime_set:=E_ExTime.eWater, setTime:=stProdParam.stRecipe.ExpirationTime_Water);
END_IF


(*
IF stProdParam.eStatus=E_Prod_Status.Active 
AND refElement.State>=E_Element_State_Long.eWaterReady
THEN;
	IF refElement.memoDissolving_active 
	//OR eStatus>=E_Element_State_Long.eReady
	THEN
		refElement.ExpirationTime:=stProdParam.stRecipe.ExpirationTime;
	ELSE;
		refElement.ExpirationTime:=stProdParam.stRecipe.ExpirationTime_Water;
	END_IF
	
ELSE;
	refElement.ExpirationTime:=ExDuration_Default;
END_IF
*)
END_ACTION

ACTION act_Filling:


IF TRUE 
AND bReady
AND refElement.eState_Long=E_Element_State_Long.eProduction
AND TRUE
AND TRUE
THEN;
	CASE pFilling_State OF 
		E_Filling_State.eNot_Ready:;
				pFilling_State:=E_Filling_State.eReady_ToFill;
				
		E_Filling_State.eReady_ToFill:;
				//
		E_Filling_State.eFilling_InProcess:;
				//
		
	END_CASE
ELSE;
	pFilling_State:=E_Filling_State.eNot_Ready;
END_IF

refElement.pFilling_State:=pFilling_State;

(*
IF fbInterConnection_ProL.bActive THEN;
	IF trn_Tank_Marinade THEN;
		fbElement[E_Element_List.eLine_Marinada].pFilling_State:=pFilling_State;
	ELSIF trn_Tank_Color THEN;
		fbElement[E_Element_List.eLine_Color].pFilling_State:=pFilling_State;
	END_IF	
END_IF
*)
END_ACTION

ACTION act_GetReference:
m_Set_SFCFlags_Reference();
refElement REF= fbElement[eElementID];
refState_Long REF= fbElement[eElementID].eState_Long;
//stPis_FillWater REF= stPis[valFillWater];
//stPis_FillWaterDrain REF= stPis[valFillWaterDrain];
//stPis_DrainTapWater REF= stPis[valDrainTapWater];

ref_fbTankSensors REF= g_Data.arrTanksSens[eTank_Name];
stTank_Level:=ref_fbTankSensors.get_stTankLevel();
fbTarget.set_TankLevel(set_stTankLevel:=stTank_Level);

stPis_CWIn REF= stPis[valCW_In];
stPis_CWOut	 REF= stPis[valCW_Out];

eStatus:=refState_Long;

//bRunCIP :=g_Data.b_CIP_Run;
bRunCIP := g_Data.fbElement[eElementID].m_Get_InterConnection() = E_InterConnection.ConnToCIP;
(*
stPis_Outlet		REF= g_Piston.stPis[valOutlet];
stPis_Line			REF= g_Piston.stPis[valOutlet];
stPis_TriBlender	REF= g_Piston.stPis[valOutlet];
stPis_Drain			REF= g_Piston.stPis[valOutlet];
stPis_CIP			REF= g_Piston.stPis[valOutlet];
*)
END_ACTION

ACTION act_Oper:
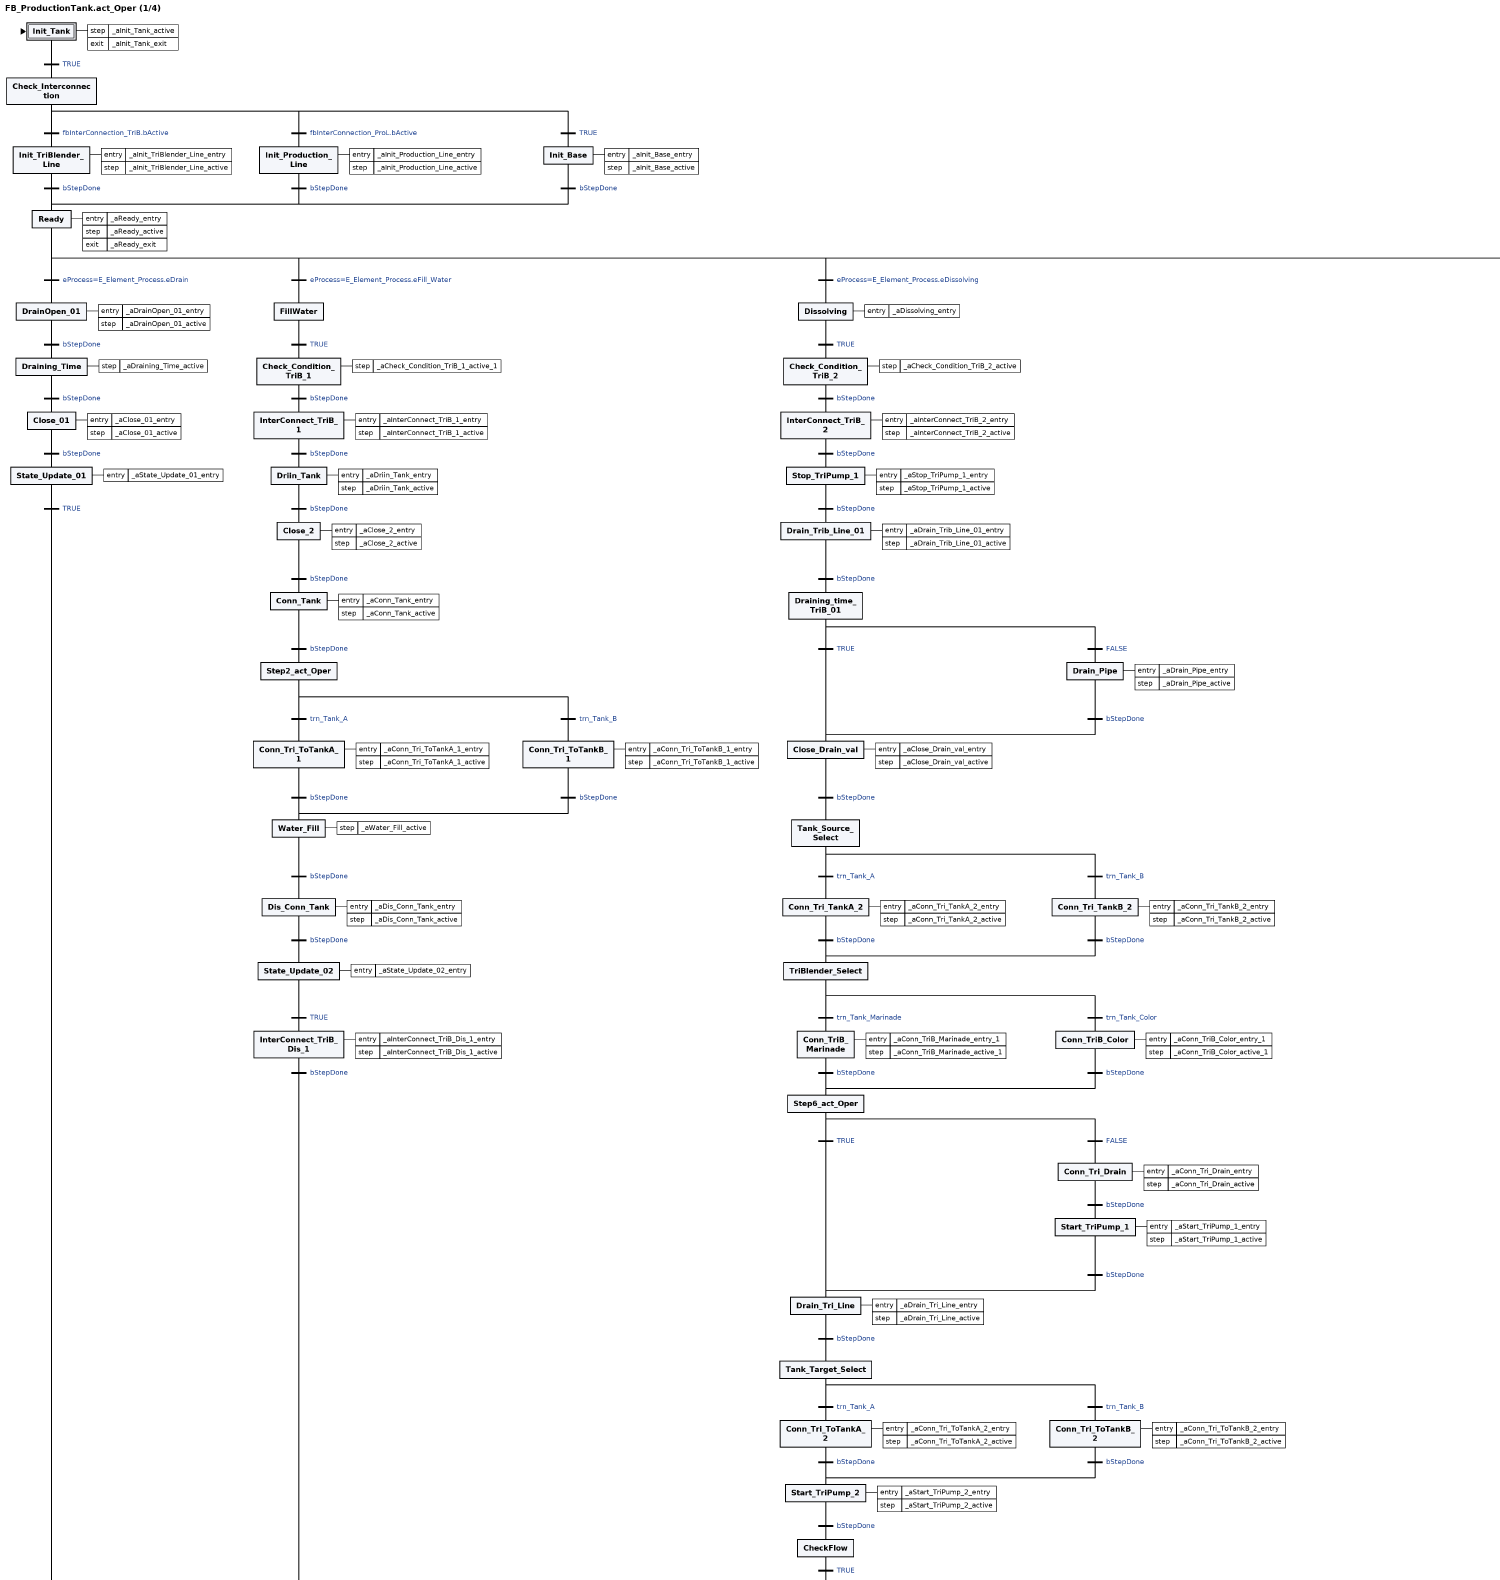
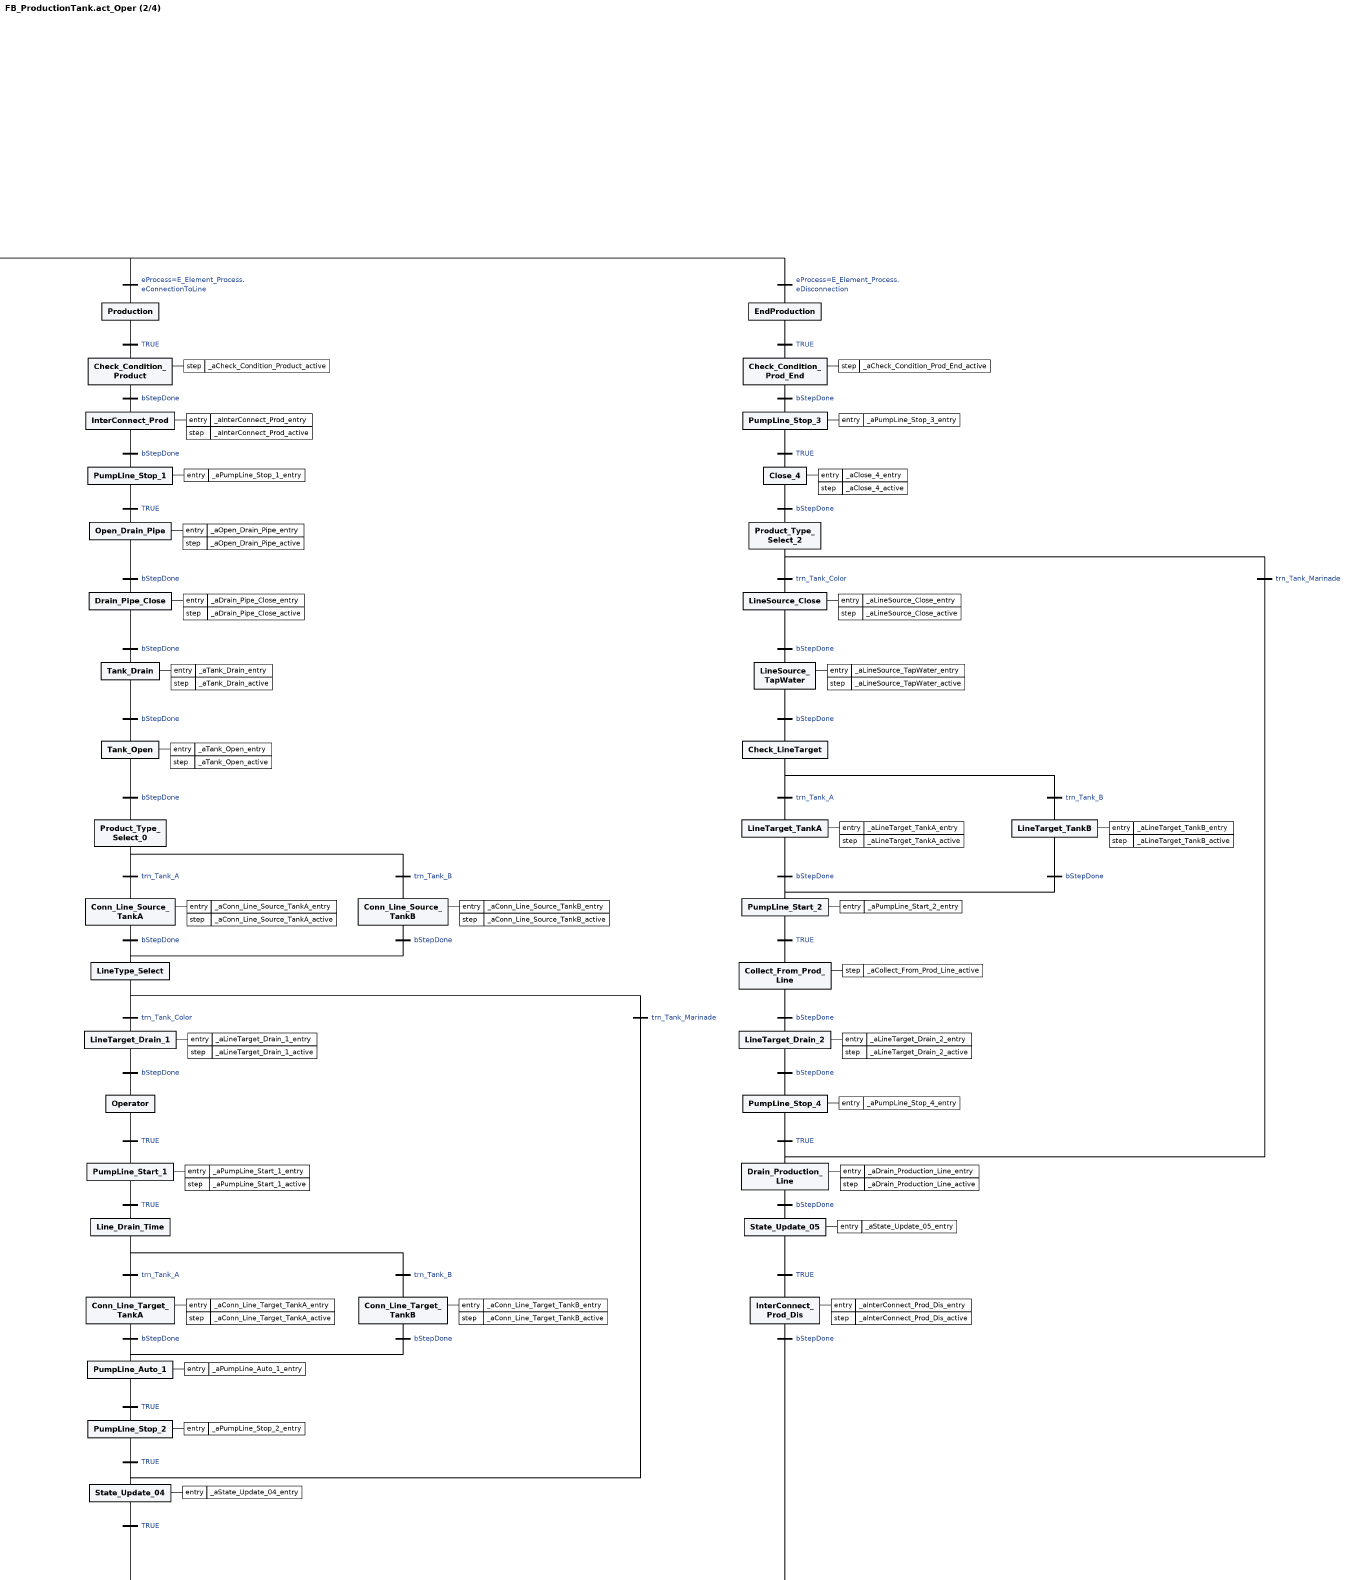
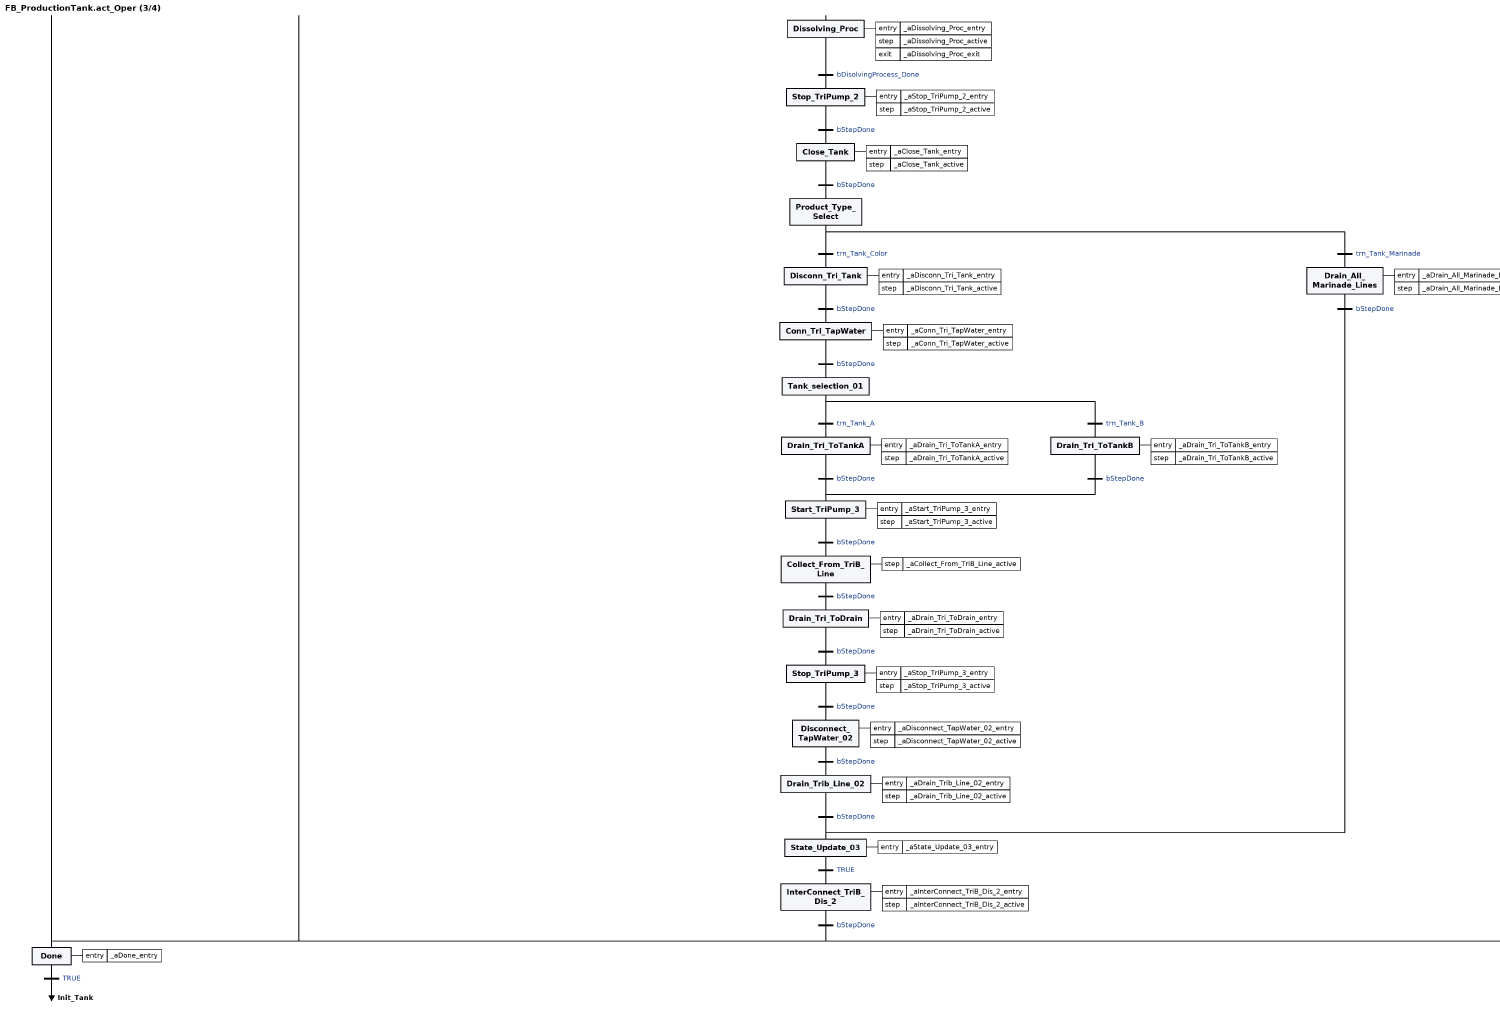
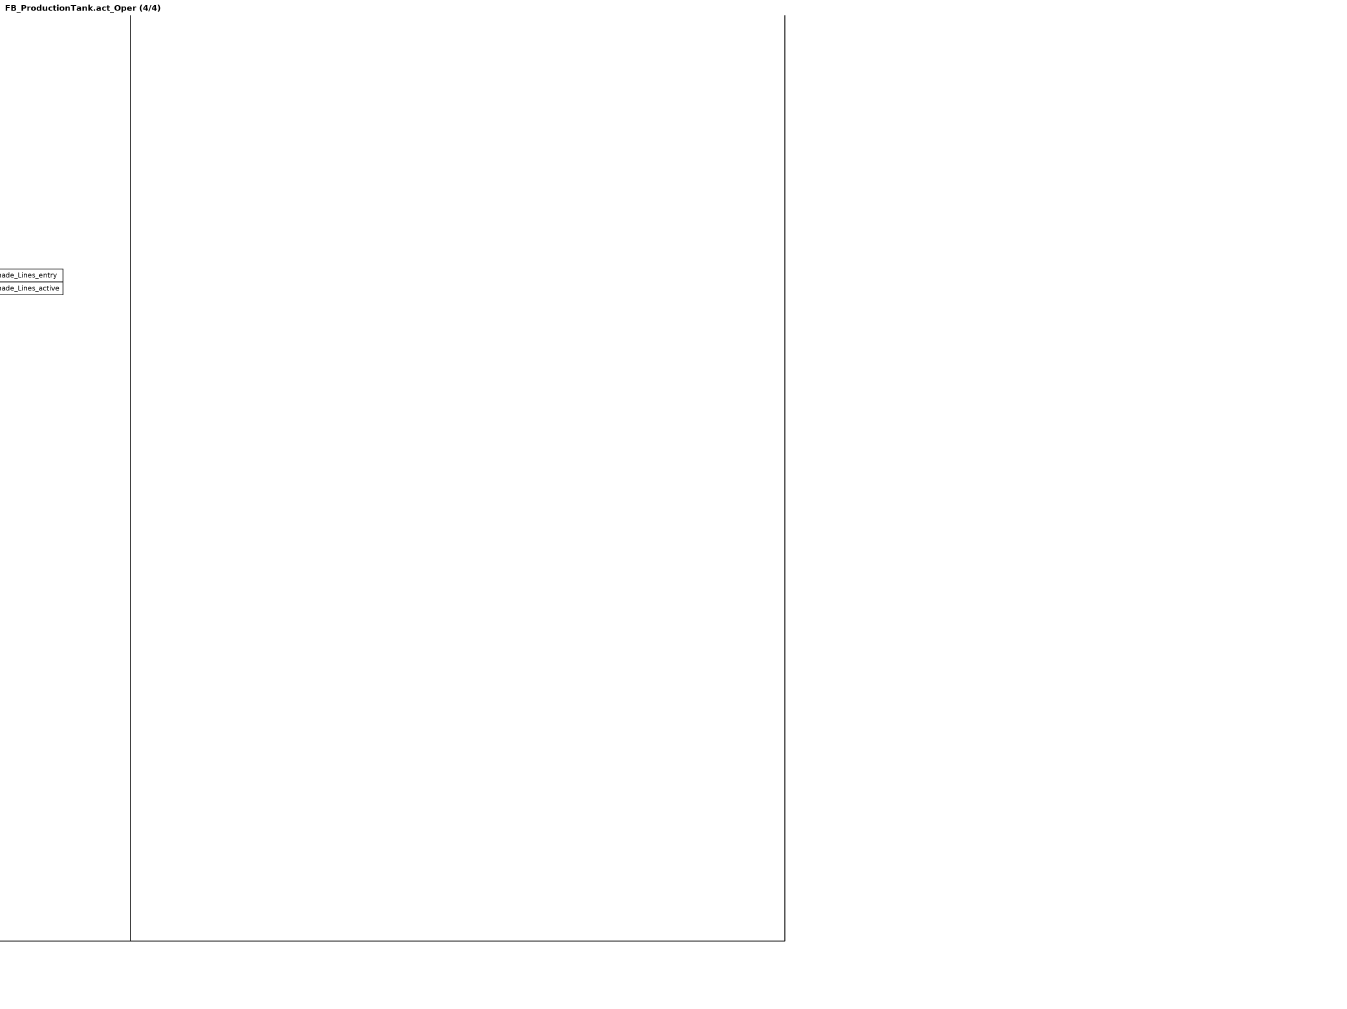
INITIAL_STEP Init_Tank:
    _aInit_Tank_active(N);  // step action
    _aInit_Tank_exit(P0);  // exit action
END_STEP
TRANSITION FROM Init_Tank TO Check_Interconnection
    := TRUE;
END_TRANSITION
STEP Check_Interconnection:
END_STEP
TRANSITION FROM Check_Interconnection TO Init_TriBlender_Line
    := fbInterConnection_TriB.bActive;
END_TRANSITION
STEP Init_TriBlender_Line:
    _aInit_TriBlender_Line_entry(P1);  // entry action
    _aInit_TriBlender_Line_active(N);  // step action
END_STEP
TRANSITION FROM Init_TriBlender_Line TO Ready
    := bStepDone;
END_TRANSITION
TRANSITION FROM Check_Interconnection TO Init_Production_Line
    := fbInterConnection_ProL.bActive;
END_TRANSITION
STEP Init_Production_Line:
    _aInit_Production_Line_entry(P1);  // entry action
    _aInit_Production_Line_active(N);  // step action
END_STEP
TRANSITION FROM Init_Production_Line TO Ready
    := bStepDone;
END_TRANSITION
TRANSITION FROM Check_Interconnection TO Init_Base
    := TRUE;
END_TRANSITION
STEP Init_Base:
    _aInit_Base_entry(P1);  // entry action
    _aInit_Base_active(N);  // step action
END_STEP
TRANSITION FROM Init_Base TO Ready
    := bStepDone;
END_TRANSITION
STEP Ready:
    _aReady_entry(P1);  // entry action
    _aReady_active(N);  // step action
    _aReady_exit(P0);  // exit action
END_STEP
TRANSITION FROM Ready TO DrainOpen_01
    := eProcess=E_Element_Process.eDrain;
END_TRANSITION
STEP DrainOpen_01:  // min time T#2s
    _aDrainOpen_01_entry(P1);  // entry action
    _aDrainOpen_01_active(N);  // step action
END_STEP
TRANSITION FROM DrainOpen_01 TO Draining_Time
    := bStepDone;
END_TRANSITION
STEP Draining_Time:  // min time T#2s
    _aDraining_Time_active(N);  // step action
END_STEP
TRANSITION FROM Draining_Time TO Close_01
    := bStepDone;
END_TRANSITION
STEP Close_01:  // min time T#2s
    _aClose_01_entry(P1);  // entry action
    _aClose_01_active(N);  // step action
END_STEP
TRANSITION FROM Close_01 TO State_Update_01
    := bStepDone;
END_TRANSITION
STEP State_Update_01:
    _aState_Update_01_entry(P1);  // entry action
END_STEP
TRANSITION FROM State_Update_01 TO Done
    := TRUE;
END_TRANSITION
TRANSITION FROM Ready TO FillWater
    := eProcess=E_Element_Process.eFill_Water;
END_TRANSITION
STEP FillWater:
END_STEP
TRANSITION FROM FillWater TO Check_Condition_TriB_1
    := TRUE;
END_TRANSITION
STEP Check_Condition_TriB_1:
    _aCheck_Condition_TriB_1_active_1(N);  // step action
END_STEP
TRANSITION FROM Check_Condition_TriB_1 TO InterConnect_TriB_1
    := bStepDone;
END_TRANSITION
STEP InterConnect_TriB_1:
    _aInterConnect_TriB_1_entry(P1);  // entry action
    _aInterConnect_TriB_1_active(N);  // step action
END_STEP
TRANSITION FROM InterConnect_TriB_1 TO Driin_Tank
    := bStepDone;
END_TRANSITION
STEP Driin_Tank:  // min time t#2s
    _aDriin_Tank_entry(P1);  // entry action
    _aDriin_Tank_active(N);  // step action
END_STEP
TRANSITION FROM Driin_Tank TO Close_2
    := bStepDone;
END_TRANSITION
STEP Close_2:  // min time t#2s
    _aClose_2_entry(P1);  // entry action
    _aClose_2_active(N);  // step action
END_STEP
TRANSITION FROM Close_2 TO Conn_Tank
    := bStepDone;
END_TRANSITION
STEP Conn_Tank:  // min time t#2s
    _aConn_Tank_entry(P1);  // entry action
    _aConn_Tank_active(N);  // step action
END_STEP
TRANSITION FROM Conn_Tank TO Step2_act_Oper
    := bStepDone;
END_TRANSITION
STEP Step2_act_Oper:
END_STEP
TRANSITION FROM Step2_act_Oper TO Conn_Tri_ToTankA_1
    := trn_Tank_A;
END_TRANSITION
STEP Conn_Tri_ToTankA_1:
    _aConn_Tri_ToTankA_1_entry(P1);  // entry action
    _aConn_Tri_ToTankA_1_active(N);  // step action
END_STEP
TRANSITION FROM Conn_Tri_ToTankA_1 TO Water_Fill
    := bStepDone;
END_TRANSITION
TRANSITION FROM Step2_act_Oper TO Conn_Tri_ToTankB_1
    := trn_Tank_B;
END_TRANSITION
STEP Conn_Tri_ToTankB_1:
    _aConn_Tri_ToTankB_1_entry(P1);  // entry action
    _aConn_Tri_ToTankB_1_active(N);  // step action
END_STEP
TRANSITION FROM Conn_Tri_ToTankB_1 TO Water_Fill
    := bStepDone;
END_TRANSITION
STEP Water_Fill:  // min time t#2s
    _aWater_Fill_active(N);  // step action
END_STEP
TRANSITION FROM Water_Fill TO Dis_Conn_Tank
    := bStepDone;
END_TRANSITION
STEP Dis_Conn_Tank:  // min time t#2s
    _aDis_Conn_Tank_entry(P1);  // entry action
    _aDis_Conn_Tank_active(N);  // step action
END_STEP
TRANSITION FROM Dis_Conn_Tank TO State_Update_02
    := bStepDone;
END_TRANSITION
STEP State_Update_02:  // min time t#2s
    _aState_Update_02_entry(P1);  // entry action
END_STEP
TRANSITION FROM State_Update_02 TO InterConnect_TriB_Dis_1
    := TRUE;
END_TRANSITION
STEP InterConnect_TriB_Dis_1:
    _aInterConnect_TriB_Dis_1_entry(P1);  // entry action
    _aInterConnect_TriB_Dis_1_active(N);  // step action
END_STEP
TRANSITION FROM InterConnect_TriB_Dis_1 TO Done
    := bStepDone;
END_TRANSITION
TRANSITION FROM Ready TO Dissolving
    := eProcess=E_Element_Process.eDissolving;
END_TRANSITION
STEP Dissolving:
    _aDissolving_entry(P1);  // entry action
END_STEP
TRANSITION FROM Dissolving TO Check_Condition_TriB_2
    := TRUE;
END_TRANSITION
STEP Check_Condition_TriB_2:
    _aCheck_Condition_TriB_2_active(N);  // step action
END_STEP
TRANSITION FROM Check_Condition_TriB_2 TO InterConnect_TriB_2
    := bStepDone;
END_TRANSITION
STEP InterConnect_TriB_2:
    _aInterConnect_TriB_2_entry(P1);  // entry action
    _aInterConnect_TriB_2_active(N);  // step action
END_STEP
TRANSITION FROM InterConnect_TriB_2 TO Stop_TriPump_1
    := bStepDone;
END_TRANSITION
STEP Stop_TriPump_1:
    _aStop_TriPump_1_entry(P1);  // entry action
    _aStop_TriPump_1_active(N);  // step action
END_STEP
TRANSITION FROM Stop_TriPump_1 TO Drain_Trib_Line_01
    := bStepDone;
END_TRANSITION
STEP Drain_Trib_Line_01:
    _aDrain_Trib_Line_01_entry(P1);  // entry action
    _aDrain_Trib_Line_01_active(N);  // step action
END_STEP
TRANSITION FROM Drain_Trib_Line_01 TO Draining_time_TriB_01
    := bStepDone;
END_TRANSITION
STEP Draining_time_TriB_01:  // min time T#10s
END_STEP
TRANSITION FROM Draining_time_TriB_01 TO Close_Drain_val
    := TRUE;
END_TRANSITION
TRANSITION FROM Draining_time_TriB_01 TO Drain_Pipe
    := FALSE;
END_TRANSITION
STEP Drain_Pipe:  // min time T#2s
    _aDrain_Pipe_entry(P1);  // entry action
    _aDrain_Pipe_active(N);  // step action
END_STEP
TRANSITION FROM Drain_Pipe TO Close_Drain_val
    := bStepDone;
END_TRANSITION
STEP Close_Drain_val:
    _aClose_Drain_val_entry(P1);  // entry action
    _aClose_Drain_val_active(N);  // step action
END_STEP
TRANSITION FROM Close_Drain_val TO Tank_Source_Select
    := bStepDone;
END_TRANSITION
STEP Tank_Source_Select:
END_STEP
TRANSITION FROM Tank_Source_Select TO Conn_Tri_TankA_2
    := trn_Tank_A;
END_TRANSITION
STEP Conn_Tri_TankA_2:
    _aConn_Tri_TankA_2_entry(P1);  // entry action
    _aConn_Tri_TankA_2_active(N);  // step action
END_STEP
TRANSITION FROM Conn_Tri_TankA_2 TO TriBlender_Select
    := bStepDone;
END_TRANSITION
TRANSITION FROM Tank_Source_Select TO Conn_Tri_TankB_2
    := trn_Tank_B;
END_TRANSITION
STEP Conn_Tri_TankB_2:
    _aConn_Tri_TankB_2_entry(P1);  // entry action
    _aConn_Tri_TankB_2_active(N);  // step action
END_STEP
TRANSITION FROM Conn_Tri_TankB_2 TO TriBlender_Select
    := bStepDone;
END_TRANSITION
STEP TriBlender_Select:
END_STEP
TRANSITION FROM TriBlender_Select TO Conn_TriB_Marinade
    := trn_Tank_Marinade;
END_TRANSITION
STEP Conn_TriB_Marinade:
    _aConn_TriB_Marinade_entry_1(P1);  // entry action
    _aConn_TriB_Marinade_active_1(N);  // step action
END_STEP
TRANSITION FROM Conn_TriB_Marinade TO Step6_act_Oper
    := bStepDone;
END_TRANSITION
TRANSITION FROM TriBlender_Select TO Conn_TriB_Color
    := trn_Tank_Color;
END_TRANSITION
STEP Conn_TriB_Color:
    _aConn_TriB_Color_entry_1(P1);  // entry action
    _aConn_TriB_Color_active_1(N);  // step action
END_STEP
TRANSITION FROM Conn_TriB_Color TO Step6_act_Oper
    := bStepDone;
END_TRANSITION
STEP Step6_act_Oper:
END_STEP
TRANSITION FROM Step6_act_Oper TO Drain_Tri_Line
    := TRUE;
END_TRANSITION
TRANSITION FROM Step6_act_Oper TO Conn_Tri_Drain
    := FALSE;
END_TRANSITION
STEP Conn_Tri_Drain:
    _aConn_Tri_Drain_entry(P1);  // entry action
    _aConn_Tri_Drain_active(N);  // step action
END_STEP
TRANSITION FROM Conn_Tri_Drain TO Start_TriPump_1
    := bStepDone;
END_TRANSITION
STEP Start_TriPump_1:
    _aStart_TriPump_1_entry(P1);  // entry action
    _aStart_TriPump_1_active(N);  // step action
END_STEP
TRANSITION FROM Start_TriPump_1 TO Drain_Tri_Line
    := bStepDone;
END_TRANSITION
STEP Drain_Tri_Line:  // min time T#10s
    _aDrain_Tri_Line_entry(P1);  // entry action
    _aDrain_Tri_Line_active(N);  // step action
END_STEP
TRANSITION FROM Drain_Tri_Line TO Tank_Target_Select
    := bStepDone;
END_TRANSITION
STEP Tank_Target_Select:
END_STEP
TRANSITION FROM Tank_Target_Select TO Conn_Tri_ToTankA_2
    := trn_Tank_A;
END_TRANSITION
STEP Conn_Tri_ToTankA_2:
    _aConn_Tri_ToTankA_2_entry(P1);  // entry action
    _aConn_Tri_ToTankA_2_active(N);  // step action
END_STEP
TRANSITION FROM Conn_Tri_ToTankA_2 TO Start_TriPump_2
    := bStepDone;
END_TRANSITION
TRANSITION FROM Tank_Target_Select TO Conn_Tri_ToTankB_2
    := trn_Tank_B;
END_TRANSITION
STEP Conn_Tri_ToTankB_2:
    _aConn_Tri_ToTankB_2_entry(P1);  // entry action
    _aConn_Tri_ToTankB_2_active(N);  // step action
END_STEP
TRANSITION FROM Conn_Tri_ToTankB_2 TO Start_TriPump_2
    := bStepDone;
END_TRANSITION
STEP Start_TriPump_2:
    _aStart_TriPump_2_entry(P1);  // entry action
    _aStart_TriPump_2_active(N);  // step action
END_STEP
TRANSITION FROM Start_TriPump_2 TO CheckFlow
    := bStepDone;
END_TRANSITION
STEP CheckFlow:  // min time t#20s
END_STEP
TRANSITION FROM CheckFlow TO Dissolving_Proc
    := TRUE;
END_TRANSITION
STEP Dissolving_Proc:
    _aDissolving_Proc_entry(P1);  // entry action
    _aDissolving_Proc_active(N);  // step action
    _aDissolving_Proc_exit(P0);  // exit action
END_STEP
TRANSITION FROM Dissolving_Proc TO Stop_TriPump_2
    := bDisolvingProcess_Done;
END_TRANSITION
STEP Stop_TriPump_2:  // min time T#5s
    _aStop_TriPump_2_entry(P1);  // entry action
    _aStop_TriPump_2_active(N);  // step action
END_STEP
TRANSITION FROM Stop_TriPump_2 TO Close_Tank
    := bStepDone;
END_TRANSITION
STEP Close_Tank:
    _aClose_Tank_entry(P1);  // entry action
    _aClose_Tank_active(N);  // step action
END_STEP
TRANSITION FROM Close_Tank TO Product_Type_Select
    := bStepDone;
END_TRANSITION
STEP Product_Type_Select:
END_STEP
TRANSITION FROM Product_Type_Select TO Disconn_Tri_Tank
    := trn_Tank_Color;
END_TRANSITION
STEP Disconn_Tri_Tank:  // min time t#100ms
    _aDisconn_Tri_Tank_entry(P1);  // entry action
    _aDisconn_Tri_Tank_active(N);  // step action
END_STEP
TRANSITION FROM Disconn_Tri_Tank TO Conn_Tri_TapWater
    := bStepDone;
END_TRANSITION
STEP Conn_Tri_TapWater:  // min time T#5s
    _aConn_Tri_TapWater_entry(P1);  // entry action
    _aConn_Tri_TapWater_active(N);  // step action
END_STEP
TRANSITION FROM Conn_Tri_TapWater TO Tank_selection_01
    := bStepDone;
END_TRANSITION
STEP Tank_selection_01:
END_STEP
TRANSITION FROM Tank_selection_01 TO Drain_Tri_ToTankA
    := trn_Tank_A;
END_TRANSITION
STEP Drain_Tri_ToTankA:  // min time t#100ms
    _aDrain_Tri_ToTankA_entry(P1);  // entry action
    _aDrain_Tri_ToTankA_active(N);  // step action
END_STEP
TRANSITION FROM Drain_Tri_ToTankA TO Start_TriPump_3
    := bStepDone;
END_TRANSITION
TRANSITION FROM Tank_selection_01 TO Drain_Tri_ToTankB
    := trn_Tank_B;
END_TRANSITION
STEP Drain_Tri_ToTankB:  // min time t#100ms
    _aDrain_Tri_ToTankB_entry(P1);  // entry action
    _aDrain_Tri_ToTankB_active(N);  // step action
END_STEP
TRANSITION FROM Drain_Tri_ToTankB TO Start_TriPump_3
    := bStepDone;
END_TRANSITION
STEP Start_TriPump_3:
    _aStart_TriPump_3_entry(P1);  // entry action
    _aStart_TriPump_3_active(N);  // step action
END_STEP
TRANSITION FROM Start_TriPump_3 TO Collect_From_TriB_Line
    := bStepDone;
END_TRANSITION
STEP Collect_From_TriB_Line:
    _aCollect_From_TriB_Line_active(N);  // step action
END_STEP
TRANSITION FROM Collect_From_TriB_Line TO Drain_Tri_ToDrain
    := bStepDone;
END_TRANSITION
STEP Drain_Tri_ToDrain:  // min time T#25s
    _aDrain_Tri_ToDrain_entry(P1);  // entry action
    _aDrain_Tri_ToDrain_active(N);  // step action
END_STEP
TRANSITION FROM Drain_Tri_ToDrain TO Stop_TriPump_3
    := bStepDone;
END_TRANSITION
STEP Stop_TriPump_3:
    _aStop_TriPump_3_entry(P1);  // entry action
    _aStop_TriPump_3_active(N);  // step action
END_STEP
TRANSITION FROM Stop_TriPump_3 TO Disconnect_TapWater_02
    := bStepDone;
END_TRANSITION
STEP Disconnect_TapWater_02:
    _aDisconnect_TapWater_02_entry(P1);  // entry action
    _aDisconnect_TapWater_02_active(N);  // step action
END_STEP
TRANSITION FROM Disconnect_TapWater_02 TO Drain_Trib_Line_02
    := bStepDone;
END_TRANSITION
STEP Drain_Trib_Line_02:  // min time T#10s
    _aDrain_Trib_Line_02_entry(P1);  // entry action
    _aDrain_Trib_Line_02_active(N);  // step action
END_STEP
TRANSITION FROM Drain_Trib_Line_02 TO State_Update_03
    := bStepDone;
END_TRANSITION
TRANSITION FROM Product_Type_Select TO Drain_All_Marinade_Lines
    := trn_Tank_Marinade;
END_TRANSITION
STEP Drain_All_Marinade_Lines:
    _aDrain_All_Marinade_Lines_entry(P1);  // entry action
    _aDrain_All_Marinade_Lines_active(N);  // step action
END_STEP
TRANSITION FROM Drain_All_Marinade_Lines TO State_Update_03
    := bStepDone;
END_TRANSITION
STEP State_Update_03:
    _aState_Update_03_entry(P1);  // entry action
END_STEP
TRANSITION FROM State_Update_03 TO InterConnect_TriB_Dis_2
    := TRUE;
END_TRANSITION
STEP InterConnect_TriB_Dis_2:
    _aInterConnect_TriB_Dis_2_entry(P1);  // entry action
    _aInterConnect_TriB_Dis_2_active(N);  // step action
END_STEP
TRANSITION FROM InterConnect_TriB_Dis_2 TO Done
    := bStepDone;
END_TRANSITION
TRANSITION FROM Ready TO Production
    := eProcess=E_Element_Process.eConnectionToLine;
END_TRANSITION
STEP Production:
END_STEP
TRANSITION FROM Production TO Check_Condition_Product
    := TRUE;
END_TRANSITION
STEP Check_Condition_Product:
    _aCheck_Condition_Product_active(N);  // step action
END_STEP
TRANSITION FROM Check_Condition_Product TO InterConnect_Prod
    := bStepDone;
END_TRANSITION
STEP InterConnect_Prod:
    _aInterConnect_Prod_entry(P1);  // entry action
    _aInterConnect_Prod_active(N);  // step action
END_STEP
TRANSITION FROM InterConnect_Prod TO PumpLine_Stop_1
    := bStepDone;
END_TRANSITION
STEP PumpLine_Stop_1:
    _aPumpLine_Stop_1_entry(P1);  // entry action
END_STEP
TRANSITION FROM PumpLine_Stop_1 TO Open_Drain_Pipe
    := TRUE;
END_TRANSITION
STEP Open_Drain_Pipe:  // min time T#5s
    _aOpen_Drain_Pipe_entry(P1);  // entry action
    _aOpen_Drain_Pipe_active(N);  // step action
END_STEP
TRANSITION FROM Open_Drain_Pipe TO Drain_Pipe_Close
    := bStepDone;
END_TRANSITION
STEP Drain_Pipe_Close:
    _aDrain_Pipe_Close_entry(P1);  // entry action
    _aDrain_Pipe_Close_active(N);  // step action
END_STEP
TRANSITION FROM Drain_Pipe_Close TO Tank_Drain
    := bStepDone;
END_TRANSITION
STEP Tank_Drain:  // min time t#2s
    _aTank_Drain_entry(P1);  // entry action
    _aTank_Drain_active(N);  // step action
END_STEP
TRANSITION FROM Tank_Drain TO Tank_Open
    := bStepDone;
END_TRANSITION
STEP Tank_Open:  // min time t#2s
    _aTank_Open_entry(P1);  // entry action
    _aTank_Open_active(N);  // step action
END_STEP
TRANSITION FROM Tank_Open TO Product_Type_Select_0
    := bStepDone;
END_TRANSITION
STEP Product_Type_Select_0:
END_STEP
TRANSITION FROM Product_Type_Select_0 TO Conn_Line_Source_TankA
    := trn_Tank_A;
END_TRANSITION
STEP Conn_Line_Source_TankA:  // min time t#100ms
    _aConn_Line_Source_TankA_entry(P1);  // entry action
    _aConn_Line_Source_TankA_active(N);  // step action
END_STEP
TRANSITION FROM Conn_Line_Source_TankA TO LineType_Select
    := bStepDone;
END_TRANSITION
TRANSITION FROM Product_Type_Select_0 TO Conn_Line_Source_TankB
    := trn_Tank_B;
END_TRANSITION
STEP Conn_Line_Source_TankB:  // min time t#100ms
    _aConn_Line_Source_TankB_entry(P1);  // entry action
    _aConn_Line_Source_TankB_active(N);  // step action
END_STEP
TRANSITION FROM Conn_Line_Source_TankB TO LineType_Select
    := bStepDone;
END_TRANSITION
STEP LineType_Select:
END_STEP
TRANSITION FROM LineType_Select TO LineTarget_Drain_1
    := trn_Tank_Color;
END_TRANSITION
STEP LineTarget_Drain_1:
    _aLineTarget_Drain_1_entry(P1);  // entry action
    _aLineTarget_Drain_1_active(N);  // step action
END_STEP
TRANSITION FROM LineTarget_Drain_1 TO Operator
    := bStepDone;
END_TRANSITION
STEP Operator:
END_STEP
TRANSITION FROM Operator TO PumpLine_Start_1
    := TRUE;
END_TRANSITION
STEP PumpLine_Start_1:
    _aPumpLine_Start_1_entry(P1);  // entry action
    _aPumpLine_Start_1_active(N);  // step action
END_STEP
TRANSITION FROM PumpLine_Start_1 TO Line_Drain_Time
    := TRUE;
END_TRANSITION
STEP Line_Drain_Time:  // min time T#10s
END_STEP
TRANSITION FROM Line_Drain_Time TO Conn_Line_Target_TankA
    := trn_Tank_A;
END_TRANSITION
STEP Conn_Line_Target_TankA:
    _aConn_Line_Target_TankA_entry(P1);  // entry action
    _aConn_Line_Target_TankA_active(N);  // step action
END_STEP
TRANSITION FROM Conn_Line_Target_TankA TO PumpLine_Auto_1
    := bStepDone;
END_TRANSITION
TRANSITION FROM Line_Drain_Time TO Conn_Line_Target_TankB
    := trn_Tank_B;
END_TRANSITION
STEP Conn_Line_Target_TankB:
    _aConn_Line_Target_TankB_entry(P1);  // entry action
    _aConn_Line_Target_TankB_active(N);  // step action
END_STEP
TRANSITION FROM Conn_Line_Target_TankB TO PumpLine_Auto_1
    := bStepDone;
END_TRANSITION
STEP PumpLine_Auto_1:
    _aPumpLine_Auto_1_entry(P1);  // entry action
END_STEP
TRANSITION FROM PumpLine_Auto_1 TO PumpLine_Stop_2
    := TRUE;
END_TRANSITION
STEP PumpLine_Stop_2:
    _aPumpLine_Stop_2_entry(P1);  // entry action
END_STEP
TRANSITION FROM PumpLine_Stop_2 TO State_Update_04
    := TRUE;
END_TRANSITION
TRANSITION FROM LineType_Select TO State_Update_04
    := trn_Tank_Marinade;
END_TRANSITION
STEP State_Update_04:
    _aState_Update_04_entry(P1);  // entry action
END_STEP
TRANSITION FROM State_Update_04 TO Done
    := TRUE;
END_TRANSITION
TRANSITION FROM Ready TO EndProduction
    := eProcess=E_Element_Process.eDisconnection;
END_TRANSITION
STEP EndProduction:
END_STEP
TRANSITION FROM EndProduction TO Check_Condition_Prod_End
    := TRUE;
END_TRANSITION
STEP Check_Condition_Prod_End:
    _aCheck_Condition_Prod_End_active(N);  // step action
END_STEP
TRANSITION FROM Check_Condition_Prod_End TO PumpLine_Stop_3
    := bStepDone;
END_TRANSITION
STEP PumpLine_Stop_3:
    _aPumpLine_Stop_3_entry(P1);  // entry action
END_STEP
TRANSITION FROM PumpLine_Stop_3 TO Close_4
    := TRUE;
END_TRANSITION
STEP Close_4:
    _aClose_4_entry(P1);  // entry action
    _aClose_4_active(N);  // step action
END_STEP
TRANSITION FROM Close_4 TO Product_Type_Select_2
    := bStepDone;
END_TRANSITION
STEP Product_Type_Select_2:
END_STEP
TRANSITION FROM Product_Type_Select_2 TO LineSource_Close
    := trn_Tank_Color;
END_TRANSITION
STEP LineSource_Close:
    _aLineSource_Close_entry(P1);  // entry action
    _aLineSource_Close_active(N);  // step action
END_STEP
TRANSITION FROM LineSource_Close TO LineSource_TapWater
    := bStepDone;
END_TRANSITION
STEP LineSource_TapWater:
    _aLineSource_TapWater_entry(P1);  // entry action
    _aLineSource_TapWater_active(N);  // step action
END_STEP
TRANSITION FROM LineSource_TapWater TO Check_LineTarget
    := bStepDone;
END_TRANSITION
STEP Check_LineTarget:
END_STEP
TRANSITION FROM Check_LineTarget TO LineTarget_TankA
    := trn_Tank_A;
END_TRANSITION
STEP LineTarget_TankA:
    _aLineTarget_TankA_entry(P1);  // entry action
    _aLineTarget_TankA_active(N);  // step action
END_STEP
TRANSITION FROM LineTarget_TankA TO PumpLine_Start_2
    := bStepDone;
END_TRANSITION
TRANSITION FROM Check_LineTarget TO LineTarget_TankB
    := trn_Tank_B;
END_TRANSITION
STEP LineTarget_TankB:
    _aLineTarget_TankB_entry(P1);  // entry action
    _aLineTarget_TankB_active(N);  // step action
END_STEP
TRANSITION FROM LineTarget_TankB TO PumpLine_Start_2
    := bStepDone;
END_TRANSITION
STEP PumpLine_Start_2:
    _aPumpLine_Start_2_entry(P1);  // entry action
END_STEP
TRANSITION FROM PumpLine_Start_2 TO Collect_From_Prod_Line
    := TRUE;
END_TRANSITION
STEP Collect_From_Prod_Line:
    _aCollect_From_Prod_Line_active(N);  // step action
END_STEP
TRANSITION FROM Collect_From_Prod_Line TO LineTarget_Drain_2
    := bStepDone;
END_TRANSITION
STEP LineTarget_Drain_2:  // min time T#25s
    _aLineTarget_Drain_2_entry(P1);  // entry action
    _aLineTarget_Drain_2_active(N);  // step action
END_STEP
TRANSITION FROM LineTarget_Drain_2 TO PumpLine_Stop_4
    := bStepDone;
END_TRANSITION
STEP PumpLine_Stop_4:
    _aPumpLine_Stop_4_entry(P1);  // entry action
END_STEP
TRANSITION FROM PumpLine_Stop_4 TO Drain_Production_Line
    := TRUE;
END_TRANSITION
TRANSITION FROM Product_Type_Select_2 TO Drain_Production_Line
    := trn_Tank_Marinade;
END_TRANSITION
STEP Drain_Production_Line:
    _aDrain_Production_Line_entry(P1);  // entry action
    _aDrain_Production_Line_active(N);  // step action
END_STEP
TRANSITION FROM Drain_Production_Line TO State_Update_05
    := bStepDone;
END_TRANSITION
STEP State_Update_05:
    _aState_Update_05_entry(P1);  // entry action
END_STEP
TRANSITION FROM State_Update_05 TO InterConnect_Prod_Dis
    := TRUE;
END_TRANSITION
STEP InterConnect_Prod_Dis:
    _aInterConnect_Prod_Dis_entry(P1);  // entry action
    _aInterConnect_Prod_Dis_active(N);  // step action
END_STEP
TRANSITION FROM InterConnect_Prod_Dis TO Done
    := bStepDone;
END_TRANSITION
STEP Done:  // min time T#2s
    _aDone_entry(P1);  // entry action
END_STEP
TRANSITION FROM Done TO Init_Tank
    := TRUE;
END_TRANSITION
// branch label Branch11_act_Oper
// branch label Branch3_act_Oper
// branch label Branch10_act_Oper
// branch label Branch1_act_Oper
// branch label Branch7_act_Oper
// branch label Branch9_act_Oper
// branch label Branch2_act_Oper
// branch label Branch8_act_Oper
// branch label Branch4_act_Oper
// branch label Branch5_act_Oper
// branch label Branch14_act_Oper
// branch label Branch6_act_Oper
// branch label Branch12_act_Oper
// branch label Branch0_act_Oper_Tank
END_ACTION

ACTION act_TempCntrl:
CASE eElementID OF 
	E_Element_List.eTank_1:
		//Marinada Tank 1
		st_TempCntrl 	REF=g_ProcControl.arr_stProcCntrl[E_ProcessControl_Name.eMarinTank1_Temp];
		pc_TempCntrl 	REF= g_ProcControl.arr_fbProcCntrl[E_ProcessControl_Name.eMarinTank1_Temp];
		//tolerance
	E_Element_List.eTank_2:
		//Marinada Tank 2
		st_TempCntrl 	REF=g_ProcControl.arr_stProcCntrl[E_ProcessControl_Name.eMarinTank2_Temp];
		pc_TempCntrl 	REF= g_ProcControl.arr_fbProcCntrl[E_ProcessControl_Name.eMarinTank2_Temp];
	E_Element_List.eTank_3:
		//Color Tank 1
		st_TempCntrl 	REF=g_ProcControl.arr_stProcCntrl[E_ProcessControl_Name.eColorTank1_Temp];
		pc_TempCntrl 	REF= g_ProcControl.arr_fbProcCntrl[E_ProcessControl_Name.eColorTank1_Temp];
	E_Element_List.eTank_4:
		//Color Tank 2
		st_TempCntrl 	REF=g_ProcControl.arr_stProcCntrl[E_ProcessControl_Name.eColorTank2_Temp];
		pc_TempCntrl 	REF= g_ProcControl.arr_fbProcCntrl[E_ProcessControl_Name.eColorTank2_Temp];
END_CASE
st_TempCntrl.rValue:=g_AnalogSensor.stAnalogSensor[sens_TankTemp].Value;//sensor
//st_TempCntrl.rValue:=rTest;//sensor test
st_TempCntrl.rSetPoint:=stProdParam.stRecipe.Temperature;//value from recipe
st_TempCntrl.fHystLow:=stProdParam.stRecipe.Temperature-1;
st_TempCntrl.fHystHigh:=stProdParam.stRecipe.Temperature+0.5;
//st_TempCntrl.ToleranceHigh:=5;
//st_TempCntrl.ToleravceLow:=-55;



bCntrlTemp:=stProdParam.eStatus=E_Prod_Status.Active
AND eStatus>=E_Element_State_Long.eWaterReady;

IF bCntrlTemp AND NOT bRunCIP THEN
	//pc_TempCntrl.mRun_Hyst();
	pc_TempCntrl(stProcessControl:=st_TempCntrl);
	
 	IF TRUE 
	AND (NOT st_TempCntrl.bHystOut)
	AND  stPis_CWOut.st_Close
	THEN
		stPis_CWOut.req_Open:=TRUE;
		
	ELSIF (st_TempCntrl.bHystOut)
	AND stPis_CWOut.st_Open THEN;
		stPis_CWOut.req_Close:=TRUE;
		
	END_IF
		
	IF NOT stPis_CWIn.st_Open THEN
		stPis_CWIn.req_Open:=TRUE;
	END_IF
	
ELSE
	IF NOT stPis_CWOut.st_Close THEN;
		stPis_CWOut.req_Close:=TRUE;
	END_IF
	
	IF NOT stPis_CWIn.st_Close THEN
		stPis_CWIn.req_Close:=TRUE;
	END_IF
END_IF
END_ACTION

PROPERTY cip_Pump_linked : BOOL
GET
cip_Pump_linked:=memo_CIP_Pump_linked;
END_GET
SET
memo_CIP_Pump_linked:=cip_Pump_linked;
END_SET
END_PROPERTY

METHOD m_Get_TriBlender_Clean : BOOL
VAR_INPUT
END_VAR
CASE eElementID OF
	E_Element_List.eTank_1,E_Element_List.eTank_2:;
		m_Get_TriBlender_Clean:=fbElement[E_Element_List.eTriBlender_Color].m_Get_State_Short()=E_Element_State_Short.eClean;
	E_Element_List.eTank_3,E_Element_List.eTank_4:;
		m_Get_TriBlender_Clean:=fbElement[E_Element_List.eTriBlender_Marinada].m_Get_State_Short()=E_Element_State_Short.eClean;
	
ELSE;
	m_Get_TriBlender_Clean:=FALSE;
END_CASE
END_METHOD

METHOD m_HMI : BOOL
VAR_INPUT
END_VAR
fbEvent_echo();
event_state_Update_sum:= TO_INT(eStatus) + TO_INT(stProdParam.eStatus) + TO_INT(eProcess);

IF event_state_Update_sum_last<>event_state_Update_sum THEN;
	event_state_Update_sum_last:=event_state_Update_sum;
	fbEvent_echo.event();
END_IF

event_state_Update:=fbEvent_echo.echo;
END_METHOD

METHOD m_Production_Run_Pump : BOOL
VAR_INPUT
END_VAR
CASE stProdParam.stRecipe.eFilling_Mode OF
	E_Filling_Mode.Line_Cyrculation,
	E_Filling_Mode.Bin_Cyrculation:;	
			IF TRUE
			AND trn_Tank_Color
			AND (refState_Long=E_Element_State_Long.eProduction
				OR (refState_Long=E_Element_State_Long.eExpired 
					AND refElement.eState_Long_Expiered =E_Element_State_Long.eProduction)
			AND fbTarget.m_CheckStatus(eReqStatus:=E_Tank_Target.eOpen)) 
			AND ((trn_Tank_A 
				AND fbLineSource.m_CheckStatus(eReqStatus:=E_Line_Source.eTank_A) 
				AND fbLineTarget.m_CheckStatus(eReqStatus:=E_Line_Target.eTank_A))
					OR
				(trn_Tank_B 
				AND fbLineSource.m_CheckStatus(eReqStatus:=E_Line_Source.eTank_B) 
				AND fbLineTarget.m_CheckStatus(eReqStatus:=E_Line_Target.eTank_B)))		
			AND fbInterConnection_ProL.bActive
			AND TRUE
			THEN;
				m_Production_Run_Pump:=TRUE;
			ELSE;
				m_Production_Run_Pump:=FALSE;
			END_IF	
	E_Filling_Mode.Bin:;
				m_Production_Run_Pump:=fbFilling.pumpFilling;
				
	E_Filling_Mode.Not_Selected:;
	
END_CASE
END_METHOD

METHOD m_Set_SFCFlags_Reference : BOOL
//Set reference to SFC flags

refSFC.SFCInit REF= SFCInit;
refSFC.SFCReset REF= SFCReset;
refSFC.SFCError REF= SFCError;
refSFC.SFCEnableLimit REF= SFCEnableLimit;
refSFC.SFCErrorStep REF= SFCErrorStep;
refSFC.SFCErrorPOU REF= SFCErrorPOU;
refSFC.SFCQuitError REF= SFCQuitError;
refSFC.SFCPause REF= SFCPause;
refSFC.SFCTrans REF= SFCTrans;
refSFC.SFCCurrentStep REF= SFCCurrentStep;
refSFC.SFCTip REF= SFCTip;
refSFC.SFCTipMode REF= SFCTipMode;

// Cycle handle for SFC
m_SFC_Handle();
END_METHOD

METHOD m_Stirrer : BOOL
VAR_INPUT
END_VAR
IF eStatus>=E_Element_State_Long.eWaterReady THEN;
	IF stProdParam.eStatus=E_Prod_Status.Active THEN;
		IF fbInterConnection_TriB.bActive THEN;
			m_Stirrer_run(param:=stProdParam.stRecipe.StirrerDissolving);
		ELSIF fbInterConnection_ProL.bActive THEN;
			IF memo_Production_Storage_Mode THEN;
				m_Stirrer_run(param:=stProdParam.stRecipe.StirrerStorage);
			ELSE;
				m_Stirrer_run(param:=stProdParam.stRecipe.StirrerProduction);
			END_IF	
		ELSE;		
			m_Stirrer_run(param:=stProdParam.stRecipe.StirrerStorage);//fb_Stirrer.m_Run(RPM:=1203);
		END_IF
	ELSE;
		fb_Stirrer.m_Run(RPM:=stProdParam.stRecipe.StirrerStorage.Speed);
	END_IF
ELSIF eStatus<E_Element_State_Long.eWaterReady
AND refElement.m_Get_InterConnection()=E_InterConnection.ConnToCIP THEN;
	// controled by CIP
	m_Stirrer_run_CIP();
ELSE;
	fb_Stirrer.m_Stop();
END_IF
END_METHOD

METHOD m_Stirrer_run : BOOL
VAR_INPUT
	param: ST_Prod_Param_Stirrer;
END_VAR

VAR
	time_on: TIME;
	time_off: TIME;
	time_cycle: TIME;
	
	dint_temp: DINT;
END_VAR
dint_temp:=param.tON*60000;
time_on:=TO_TIME(dint_temp);
dint_temp:=param.tOFF*60000;
time_off:=TO_TIME(dint_temp);
time_cycle:=time_on+time_off;
tonStirrer_time(PT:=time_cycle, IN:=NOT tonStirrer_time.Q);
IF tonStirrer_time.Q THEN;
	IF bStirrerDirectionPositive THEN;
		bStirrerDirectionPositive:=FALSE;
	ELSE;
		bStirrerDirectionPositive:=TRUE;
	END_IF
END_IF
CASE param.Mode OF 
	E_Stirrer_mode.continues:;
						fb_Stirrer.m_Run(RPM:=param.Speed);
	E_Stirrer_mode.cyclic:;
					IF tonStirrer_time.ET<time_on THEN;
						IF param.Flip_mode AND trn_Tank_Marinade THEN;
							IF bStirrerDirectionPositive THEN;
								fb_Stirrer.m_Run(RPM:=param.Speed);
							ELSE;
								fb_Stirrer.m_Run(RPM:=-param.Speed);
							END_IF							
						ELSE;
							fb_Stirrer.m_Run(RPM:=param.Speed);
						END_IF
						
					ELSE
						fb_Stirrer.m_Stop();
					END_IF
	E_Stirrer_mode.off:;
						fb_Stirrer.m_Stop();
END_CASE
END_METHOD

METHOD m_Stirrer_run_CIP : BOOL
VAR_INPUT
END_VAR
IF memo_CIP_Pump_linked
AND g_Pump.fbPump[E_Pump_List.P1001].bRun
THEN;
	fb_Stirrer.m_Run(RPM:=1204);
ELSE;
	fb_Stirrer.m_Stop();
END_IF
END_METHOD

METHOD mClearProduction : BOOL
VAR_INPUT
	state: E_Element_State_Long:=E_Element_State_Long.eOff;

END_VAR

VAR
	stRecipeEmpty: ST_Prod_Recipe;
END_VAR
stProdParam.eStatus:=E_Prod_Status.Not_Active;
stProdParam.stRecipe:=stRecipeEmpty;
eReq:=E_Request_List.eNone;

IF state<>E_Element_State_Long.eOff THEN;
	refState_Long:=state;
END_IF
END_METHOD

METHOD mGet_Recipe : BOOL
VAR_INPUT
	indexRecipe: INT;

END_VAR

VAR
	i: INT;
END_VAR
IF indexRecipe <0 OR indexRecipe > g_Prod.cMax_Prod_Recipe THEN;
	RETURN;
END_IF

CASE eElementID	OF 
	E_Element_List.eTank_1,E_Element_List.eTank_2:;
		stProdParam.stRecipe:=g_Prod.arrRecipeMarinade[indexRecipe];
	E_Element_List.eTank_3,E_Element_List.eTank_4:;
  		stProdParam.stRecipe:=g_Prod.arrRecipeColor[indexRecipe];
END_CASE

FOR i:=1 TO g_Prod.cMaxCompInProduct DO
	stProdParam.arrWeightIng[i]:=stProdParam.stRecipe.arr_Component[i].rWeightPercentage/100 * stProdParam.WeightOrder;
	stProdParam.stRecipe.arr_Component[i].rWeight:=stProdParam.stRecipe.arr_Component[i].rWeightPercentage/100 * stProdParam.WeightOrder;
END_FOR
END_METHOD

METHOD mTimeProductionDuration : TIME
VAR_INPUT
END_VAR
IF dtRealTime > stProdParam.prodDT 
AND stProdParam.eStatus=E_Prod_Status.Active
THEN;
	mTimeProductionDuration:=dtRealTime - stProdParam.prodDT;
ELSE;
	mTimeProductionDuration:=T#0S;
END_IF
END_METHOD

METHOD mTimeRemainToStart : TIME
VAR_INPUT
END_VAR
IF stProdParam.eStatus=E_Prod_Status.Activation_Pending_Shift THEN;
	stProdParam.eStatus:=E_Prod_Status.Activation_Pending;
	stProdParam.prodDT:=g_Prod.dtProdTimePicker+T#2h;
END_IF


IF stProdParam.eStatus=E_Prod_Status.Activation_Pending THEN;
	IF stProdParam.prodDT > dtRealTime THEN;
		mTimeRemainToStart:=stProdParam.prodDT - dtRealTime;
	ELSIF eStatus=E_Element_State_Long.eCIP_5_Done THEN;
		stProdParam.eStatus:=E_Prod_Status.Active;
		eReq:=E_Request_List.eWaterPrepare;
	END_IF
ELSE;
	mTimeRemainToStart:=T#0S;
END_IF
END_METHOD

PROPERTY pFilling_State : E_Filling_State
GET
pFilling_State:=eFilling_State;
END_GET
SET
eFilling_State:=pFilling_State;
END_SET
END_PROPERTY

TRANSITION trn_Tank_A:
trn_Tank_A:=(eElementID=E_Element_List.eTank_1 OR eElementID=E_Element_List.eTank_3);
END_TRANSITION

TRANSITION trn_Tank_B:
trn_Tank_B:=(eElementID=E_Element_List.eTank_2 OR eElementID=E_Element_List.eTank_4);
END_TRANSITION

TRANSITION trn_Tank_Color:
trn_Tank_Color:=(eElementID=E_Element_List.eTank_3 OR eElementID=E_Element_List.eTank_4);
END_TRANSITION

TRANSITION trn_Tank_Marinade:
trn_Tank_Marinade:=(eElementID=E_Element_List.eTank_1 OR eElementID=E_Element_List.eTank_2);
END_TRANSITION

END_FUNCTION_BLOCK

(* stored: Version 1.1.0.1, ProductVersion 3.1.4024.15
   POU FB_ProductionTank: Id {7ce7ab69-2020-4b39-9932-dc5de2cb0022}, SpecialFunc None
   Folder Manage: Id {4859bb81-2525-4c2b-a781-1bdd74a1527c}
   Action _aCheck_Condition_Prod_End_active: Id {ea934447-c608-4b2d-8492-54e27aff23a1}
   Action _aCheck_Condition_Product_active: Id {5974c684-e2ea-475a-b7c0-f8bf31f474ee}
   Action _aCheck_Condition_TriB_1_active_1: Id {2514b68e-c981-4423-bfd3-97d54b3557f9}
   Action _aCheck_Condition_TriB_2_active: Id {3435a25e-e53b-4d72-86df-bdbaf94f0db9}
   Action _aClose_01_active: Id {5ab04015-c694-4f9a-9b8c-4b71239b647e}
   Action _aClose_01_entry: Id {9eeb017c-3f6d-4ecc-b10f-34b8c57ffd7e}
   Action _aClose_2_active: Id {2a994a50-9fc5-4764-a23b-9bc5372fa21a}
   Action _aClose_2_entry: Id {af8be000-2cca-431d-a649-392ef5426d55}
   Action _aClose_4_active: Id {fb27bbd8-6847-4f40-b085-f7e864fa7d84}
   Action _aClose_4_entry: Id {0dca21d9-637c-498d-acec-349d6a295729}
   Action _aClose_Drain_val_active: Id {1f8e86ab-d67f-40c0-8c33-e06ef30fd9c9}
   Action _aClose_Drain_val_entry: Id {3da53a4c-03b7-4ee1-adcf-caa5fd2148a6}
   Action _aClose_Tank_active: Id {2c06ead2-88d9-40be-895a-8f0d110ed8be}
   Action _aClose_Tank_entry: Id {5cc86289-64c2-4c76-b9c5-e140752c2508}
   Action _aCollect_From_Prod_Line_active: Id {771b979b-2440-42f1-b9e3-8aa05f11371c}
   Action _aCollect_From_TriB_Line_active: Id {5dcba99e-f46f-42f5-b819-941d4c3e4776}
   Action _aConn_Line_Source_TankA_active: Id {514f6214-c380-4464-aa57-0c01b5dc8840}
   Action _aConn_Line_Source_TankA_entry: Id {31d4d5f8-446c-43a9-8fc6-10131b5ef3a9}
   Action _aConn_Line_Source_TankB_active: Id {b18700f3-4c1a-4b2d-968b-e669679d52bc}
   Action _aConn_Line_Source_TankB_entry: Id {24ac8e3b-7815-43f6-bd47-5bf29e94d220}
   Action _aConn_Line_Target_TankA_active: Id {051bf469-ec13-4907-be90-977ce443452f}
   Action _aConn_Line_Target_TankA_entry: Id {3ed749aa-8f51-467e-8e56-e18618c5e48c}
   Action _aConn_Line_Target_TankB_active: Id {dbd5663e-c015-45b1-adb9-f851b0a02394}
   Action _aConn_Line_Target_TankB_entry: Id {3135c06b-ae22-4556-af62-d70265eee719}
   Action _aConn_Tank_active: Id {ff32bc83-3182-476f-8923-08282db126ba}
   Action _aConn_Tank_entry: Id {2f0bed0f-71b0-4f0a-b52e-3a24e43288ea}
   Action _aConn_Tri_Drain_active: Id {21e23f89-c54d-4bdb-9092-280d6a536ad3}
   Action _aConn_Tri_Drain_entry: Id {71c4c56c-665b-4d6c-b541-623bab0a3566}
   Action _aConn_Tri_TankA_2_active: Id {4364e2c0-c46b-449a-9141-25e93a2469d5}
   Action _aConn_Tri_TankA_2_entry: Id {2bd610e8-2bfa-4834-bc76-c6dfb43dde31}
   Action _aConn_Tri_TankB_2_active: Id {4ba49e8a-0ea0-4706-98b4-e821f9d70bda}
   Action _aConn_Tri_TankB_2_entry: Id {42eb9269-7614-4ba8-a4a7-1d07e283ad4c}
   Action _aConn_Tri_TapWater_active: Id {24138e04-1a15-4964-9d15-188dc29195f1}
   Action _aConn_Tri_TapWater_entry: Id {bdbd17fc-d3cd-4d43-8766-70118e5d3ab5}
   Action _aConn_Tri_ToTankA_1_active: Id {200676c2-cdec-42e8-9618-ae8ca6b9f38b}
   Action _aConn_Tri_ToTankA_1_entry: Id {0ab40394-8baf-429f-ad97-33a73351eac4}
   Action _aConn_Tri_ToTankA_2_active: Id {ffa82fd6-fba9-4843-88bc-e51623698bca}
   Action _aConn_Tri_ToTankA_2_entry: Id {3e595616-e41d-46c1-9d9d-ae530be2aedc}
   Action _aConn_Tri_ToTankB_1_active: Id {5ca0c8bb-40d6-406a-9e2c-a019061eeb07}
   Action _aConn_Tri_ToTankB_1_entry: Id {a1ddb339-c95d-4db2-9b6c-dd031cec5140}
   Action _aConn_Tri_ToTankB_2_active: Id {77f8d6f0-0a28-4bf6-bcea-6359e9a4b468}
   Action _aConn_Tri_ToTankB_2_entry: Id {5bdf7cf0-658e-4c6d-a247-741bad7443ac}
   Action _aConn_TriB_Color_active_1: Id {22686e9f-b120-4f3e-8097-7b7dd6f88ed5}
   Action _aConn_TriB_Color_entry_1: Id {820648ba-5ddc-4e60-bf03-c47dcb508deb}
   Action _aConn_TriB_Marinade_active_1: Id {f320d655-6a46-4f63-a86b-9a664d773f15}
   Action _aConn_TriB_Marinade_entry_1: Id {f9e25531-e452-47f5-8070-122aeb7239d3}
   Action _aDis_Conn_Tank_active: Id {d399ba12-cd90-4c44-8b92-acf4c24178ca}
   Action _aDis_Conn_Tank_entry: Id {9ce403e4-db3c-4066-bb85-4f28e015e1d0}
   Action _aDisconn_Tri_Tank_active: Id {4e3daae7-f788-4a9e-93f8-c893f92f4637}
   Action _aDisconn_Tri_Tank_entry: Id {08f1c6e2-9822-4dd1-8603-1c6b86dc2dc9}
   Action _aDisconnect_TapWater_02_active: Id {236a91c0-0ea2-40b4-bdfc-bc3ed6e71f6d}
   Action _aDisconnect_TapWater_02_entry: Id {9efea0c4-5d4c-401a-831f-bca9150fae6a}
   Action _aDissolving_entry: Id {a232d1b6-f4fb-4527-be1c-8a3360775849}
   Action _aDissolving_Proc_active: Id {e2eea203-140a-4f5a-bd30-6adbaa1cdec2}
   Action _aDissolving_Proc_entry: Id {28249149-8678-4a73-bb39-1576a05b85da}
   Action _aDissolving_Proc_exit: Id {eecb273b-c74f-40f2-9e29-98965fbb414e}
   Action _aDone_entry: Id {22274b2d-d139-431d-9120-18b216750139}
   Action _aDrain_All_Marinade_Lines_active: Id {899c3007-2921-4db5-938d-09f133bcad69}
   Action _aDrain_All_Marinade_Lines_entry: Id {859b2023-8ee9-4748-8df3-e36f2780d3f3}
   Action _aDrain_Pipe_active: Id {745d3851-8fef-4f4c-b40c-794f92f1f4bc}
   Action _aDrain_Pipe_Close_active: Id {50f7add1-29fd-4ffc-a42d-e7204ab16a25}
   Action _aDrain_Pipe_Close_entry: Id {07e14980-9e90-480d-84e1-53c6cf109558}
   Action _aDrain_Pipe_entry: Id {f7c9babc-9117-4ecb-8d6b-9e1ef55e0dc8}
   Action _aDrain_Production_Line_active: Id {49fa2366-38f9-4492-b91c-e1d2a1f015c6}
   Action _aDrain_Production_Line_entry: Id {9f48cf48-e395-4431-9787-264f898cfbae}
   Action _aDrain_Tri_Line_active: Id {81d134cd-a182-4f22-906b-f3879f9c0975}
   Action _aDrain_Tri_Line_entry: Id {1cbc5bf8-c1d3-405d-8d26-d1075d5f6701}
   Action _aDrain_Tri_ToDrain_active: Id {16ba7324-771a-4c87-9ee6-6423d58e799c}
   Action _aDrain_Tri_ToDrain_entry: Id {a561a662-bd87-41c2-aea4-a64ee58dffa4}
   Action _aDrain_Tri_ToTankA_active: Id {788903fd-cc72-44d4-a5cb-8bca7d2f8512}
   Action _aDrain_Tri_ToTankA_entry: Id {e6d59764-ce9a-451f-a526-36663cff2a79}
   Action _aDrain_Tri_ToTankB_active: Id {9933599e-dba5-4af5-98d0-ba1ce735c522}
   Action _aDrain_Tri_ToTankB_entry: Id {e79d7efd-5d10-44d4-9d14-f20284cfec6a}
   Action _aDrain_Trib_Line_01_active: Id {ee5a3460-3901-46e3-8704-76843715138e}
   Action _aDrain_Trib_Line_01_entry: Id {2936d130-d77f-4252-a9b7-9118c48323a5}
   Action _aDrain_Trib_Line_02_active: Id {373e0455-c3e0-4fb1-a966-aa18831efc8b}
   Action _aDrain_Trib_Line_02_entry: Id {00d2aaf8-39ef-478b-a583-a10855815d63}
   Action _aDraining_Time_active: Id {50646a45-4c33-4db3-a509-52254c9d0e39}
   Action _aDrainOpen_01_active: Id {411be806-3532-486d-8955-af87d4ed244b}
   Action _aDrainOpen_01_entry: Id {1011f731-44a1-48f7-ac02-c96fd3419d2b}
   Action _aDriin_Tank_active: Id {26ac2563-987c-433e-82de-a748503c0934}
   Action _aDriin_Tank_entry: Id {3f329f60-2c36-4d5c-a81c-6bea46c3b361}
   Action _aInit_Base_active: Id {940e813d-0beb-41d3-9670-77b30f7297d7}
   Action _aInit_Base_entry: Id {7eb9d8e6-0b86-4869-b8a2-92e36347cd42}
   Action _aInit_Production_Line_active: Id {f29a22dd-dba6-4c18-ad45-eb5a9205bc2c}
   Action _aInit_Production_Line_entry: Id {7623fe03-ad8a-4fe3-b8ee-3df8e1092a34}
   Action _aInit_Tank_active: Id {55ac947e-f328-4996-b502-0c13c5baa128}
   Action _aInit_Tank_exit: Id {cb2d02c1-4749-4191-bf76-039f0904e47d}
   Action _aInit_TriBlender_Line_active: Id {08806325-6ec1-441c-9075-35155e254ada}
   Action _aInit_TriBlender_Line_entry: Id {38b7924b-9a33-46ac-b77a-0021b8b20c00}
   Action _aInterConnect_Prod_active: Id {eb0fd1a9-b3b3-4570-b6c1-ef8289eade47}
   Action _aInterConnect_Prod_Dis_active: Id {6996a8c7-7692-424c-a264-91676cb05ae8}
   Action _aInterConnect_Prod_Dis_entry: Id {dee40ced-020e-457b-b253-7a81ce79fdc7}
   Action _aInterConnect_Prod_entry: Id {4f8e3729-9e23-4b77-841a-55532d6b8a62}
   Action _aInterConnect_TriB_1_active: Id {50aaa945-e0b8-454d-bc55-a7610b516d5c}
   Action _aInterConnect_TriB_1_entry: Id {f83eb817-3c64-4d05-91a4-e6f0efb5695f}
   Action _aInterConnect_TriB_2_active: Id {c86767af-7d54-450d-a8e4-2488e3aeaf50}
   Action _aInterConnect_TriB_2_entry: Id {c037fd38-a6e9-41af-b576-1838b786e3bb}
   Action _aInterConnect_TriB_Dis_1_active: Id {8897929d-ddfd-4a8b-91ce-9281fefd2449}
   Action _aInterConnect_TriB_Dis_1_entry: Id {f504206b-0386-428c-ab85-ea679cd1de35}
   Action _aInterConnect_TriB_Dis_2_active: Id {18799874-cd2a-4c44-9921-b705d6b002c2}
   Action _aInterConnect_TriB_Dis_2_entry: Id {922e936c-cf48-431e-91d4-f3fe0f29f04d}
   Action _aLineSource_Close_active: Id {a309b5f9-ffd7-4995-a265-4c7c8992b5f4}
   Action _aLineSource_Close_entry: Id {a03d8301-e5be-494c-aa10-2cb8828f2040}
   Action _aLineSource_TapWater_active: Id {71366205-9d33-479e-b3ed-6668795bb9be}
   Action _aLineSource_TapWater_entry: Id {ee9b6cf5-d9c5-4123-9787-9fcd70002802}
   Action _aLineTarget_Drain_1_active: Id {adb6446b-4400-4bcf-94cf-2e22730c7adb}
   Action _aLineTarget_Drain_1_entry: Id {cc014450-5112-462e-9c3c-06e7b4fbf4c6}
   Action _aLineTarget_Drain_2_active: Id {8468c3c6-0205-4718-9096-334fe5c7bc14}
   Action _aLineTarget_Drain_2_entry: Id {8a7d4cca-11e5-44ad-a00f-9c4b506ff64e}
   Action _aLineTarget_TankA_active: Id {27b3b305-7fc1-4a9e-8306-f9d32aac79a9}
   Action _aLineTarget_TankA_entry: Id {268a5449-5a38-4c9b-917e-b880df070388}
   Action _aLineTarget_TankB_active: Id {ef7ae75b-061b-40b0-b580-5003ffae5342}
   Action _aLineTarget_TankB_entry: Id {982cda96-603b-4fc8-bb44-6bd639a51537}
   Action _aOpen_Drain_Pipe_active: Id {bf201523-2d23-4f60-ba59-2a0605acfecc}
   Action _aOpen_Drain_Pipe_entry: Id {47a54e25-4d25-45d7-b66d-ae4c94120b7c}
   Action _aPumpLine_Auto_1_entry: Id {6d439a29-2ed4-43e5-8205-9d9203edcca2}
   Action _aPumpLine_Start_1_active: Id {ce6dbd88-f323-4651-bd71-86dd879d57b6}
   Action _aPumpLine_Start_1_entry: Id {dd39f47a-56ce-4e66-9fad-766c758a0414}
   Action _aPumpLine_Start_2_entry: Id {784a763c-4aaf-4759-b2cf-b5de98b7dc91}
   Action _aPumpLine_Stop_1_entry: Id {917bb24e-3637-428f-b8d1-597b829dc0e5}
   Action _aPumpLine_Stop_2_entry: Id {7e4ac8bf-96a0-48a9-849d-11f9f67b7fdc}
   Action _aPumpLine_Stop_3_entry: Id {ca23155a-4795-47b4-9628-af165468793e}
   Action _aPumpLine_Stop_4_entry: Id {792d1bb8-afca-4693-9153-1e19c39e90f9}
   Action _aReady_active: Id {86749ddf-3c7e-4ecc-9e5a-16e85de1cefc}
   Action _aReady_entry: Id {0368d597-eca6-412d-b71d-17e922d93370}
   Action _aReady_exit: Id {eda65358-fc89-414b-b675-7c61604a5bed}
   Action _aStart_TriPump_1_active: Id {e0baa26b-215d-4971-b210-61248b0a2d3a}
   Action _aStart_TriPump_1_entry: Id {eda5c941-9246-4dd3-88f8-6943eb0a83a9}
   Action _aStart_TriPump_2_active: Id {f25f79e5-4fa0-4678-b282-3b6b5431a9ae}
   Action _aStart_TriPump_2_entry: Id {f4dba2b5-c456-4682-89cb-4281e1b88ad3}
   Action _aStart_TriPump_3_active: Id {23df340a-00fb-4752-a48e-751fc143e98e}
   Action _aStart_TriPump_3_entry: Id {2651facf-f787-4997-a939-c7348845452e}
   Action _aState_Update_01_entry: Id {b174de60-7e5f-4942-be67-389d229edc22}
   Action _aState_Update_02_entry: Id {d468a8a8-6dc7-4b43-90b3-33def5e0d312}
   Action _aState_Update_03_entry: Id {4b8db616-d5f3-4549-b3e4-6ee4f44d6db0}
   Action _aState_Update_04_entry: Id {2ab0e0ff-ffd1-4ad8-87f5-e07b9ab3ae5d}
   Action _aState_Update_05_entry: Id {28f5b2ef-e541-4f70-a6c4-0fb099d990d5}
   Action _aStop_TriPump_1_active: Id {81565196-e982-4cd4-9d12-b929931661eb}
   Action _aStop_TriPump_1_entry: Id {f9c6ba37-f292-485f-a793-cd8226884d4d}
   Action _aStop_TriPump_2_active: Id {de6dd8be-1a8b-45c7-b7f8-687823dfb6aa}
   Action _aStop_TriPump_2_entry: Id {99108622-43c7-4266-b40a-522dd5604a56}
   Action _aStop_TriPump_3_active: Id {14eb9515-fba4-4878-abf3-f2c847443009}
   Action _aStop_TriPump_3_entry: Id {4c7634d9-2bc8-4efc-9c96-91473aebbd56}
   Action _aTank_Drain_active: Id {850e8108-4146-442b-badb-cf02346f4c47}
   Action _aTank_Drain_entry: Id {a299197b-3d9f-413a-9421-54b1dff00f54}
   Action _aTank_Open_active: Id {a563486c-a302-4750-9dc5-b94f9620b79e}
   Action _aTank_Open_entry: Id {540fdc51-f178-44df-9269-eb2a0262a636}
   Action _aWater_Fill_active: Id {ef2688e2-4068-4b58-bfd6-12065109d302}
   Action act_Call_Interface: Id {30d90fbf-a1e1-4624-8eba-5312c724dfd5}
   Action act_ExpirationTime: Id {232636e3-8fdc-4b48-9446-c1ccdd8dae25}
   Action act_Filling: Id {3a2f8a6e-9784-4907-89fa-be7eb4d1b7eb}
   Action act_GetReference: Id {441efe70-cf26-4ab6-bfdc-65d8c989c307}
   Action act_Oper: Id {0fa1f0eb-f194-455d-88e3-45c20b66e264}
   Action act_TempCntrl: Id {fa8d9f6d-7d99-4287-8414-2085c4b68d07}
   Property cip_Pump_linked: Id {ac226185-1e07-4925-80ab-b5fd4481a15d}
   Get Get: Id {f15d9d85-97fb-4143-b653-83a4b0989750}
   Set Set: Id {d4fd3cd6-885e-4e8b-b4a9-07e753923fb3}
   Method m_Get_TriBlender_Clean: Id {13b7f4ac-db6a-45d8-9c4a-691ded0763a9}
   Method m_HMI: Id {eaa75ffd-8860-40ef-b20b-3b03fd8650af}
   Method m_Production_Run_Pump: Id {f8a03de4-a449-4107-bdd3-bbaa65bdeb7f}
   Method m_Set_SFCFlags_Reference: Id {e572de0c-3d24-464d-bb17-5deb316affd4}
   Method m_Stirrer: Id {1b833e49-1ddd-4651-b81e-debe24950272}
   Method m_Stirrer_run: Id {307ad28f-b5d2-4fb4-8a9d-9a8b36372bf8}
   Method m_Stirrer_run_CIP: Id {c8799238-5523-43fc-a069-a2104bf79383}
   Method mClearProduction: Id {58c4c9c9-8cf2-41f1-b206-eaacde8cd18f}
   Method mGet_Recipe: Id {b8cd2ec5-ec05-4d19-a0b3-16991b77e5a1}
   Method mTimeProductionDuration: Id {b2a492d8-93d6-4df6-bd37-f2e46985a2d9}
   Method mTimeRemainToStart: Id {7d6f306c-e772-4eb3-a87e-556a8ea27eb4}
   Property pFilling_State: Id {dc44f564-aa7d-4e11-8e9c-e57e1d797297}
   Get Get: Id {21a765eb-1b41-414a-bd4e-3741aa59b706}
   Set Set: Id {2d78626e-f70c-4d07-994f-8331d9e5c207}
   Transition trn_Tank_A: Id {7f0e7518-f66a-4b4a-b16b-a3f65f501415}
   Transition trn_Tank_B: Id {e4cef271-82c6-43c9-bc0b-ff7cff0b1929}
   Transition trn_Tank_Color: Id {0f0ea737-6af2-4efd-ad50-e1b6006f4bda}
   Transition trn_Tank_Marinade: Id {706b7960-c75d-4ac2-8026-39ed0770109f} *)
